(* IEC 61131-3 sources: Antarbhukti-LLM/DatasetCreation/SeedSTs/batch1_filtered_BASIC, 119 files *)

(* ---- A_TRIG.ST ---- *)
(*@PROPERTIES_EX@
TYPE: POU
LOCALE: 0
IEC_LANGUAGE: ST
PLC_TYPE: independent
PROC_TYPE: independent
GROUP: LOGIC.GENERATORS
*)
(*@KEY@:DESCRIPTION*)
version 1.1	23. oct. 2008
programmer 	hugo
tested by	oscat

this block is similar to the IEC Standard R_trig and F_trig but it monitors a REAL for change.
if the valiue on IN changes more then D from the last value it will generate trigger and display the difference in output D.
the trigger will only be active for one cycle.
(*@KEY@:END_DESCRIPTION*)
FUNCTION_BLOCK A_TRIG

(*Group:Default*)

VAR_INPUT
	IN :	REAL;
	RES :	REAL;
END_VAR

VAR_OUTPUT
	Q :	BOOL;
	D :	REAL;
END_VAR

VAR
	last_in :	REAL;
END_VAR

(*@KEY@: WORKSHEET
NAME: A_TRIG
IEC_LANGUAGE: ST
*)
D := IN - LAST_IN;
IF ABS(D) >= res THEN
	Q := TRUE;
	last_in := IN;
ELSE
	Q := FALSE;
END_IF;

(* revision history

hm 	16. jul. 2008	rev 1.0
	original version released

hm	23. oct. 2008	rev 1.1
	code optimization
*)
(*@KEY@: END_WORKSHEET *)
END_FUNCTION_BLOCK

(* ---- AIN1.ST ---- *)
(*@PROPERTIES_EX@
TYPE: POU
LOCALE: 0
IEC_LANGUAGE: ST
PLC_TYPE: independent
PROC_TYPE: independent
GROUP: ENGINEERING.SIGNAL_PROCESSING
*)
(*@KEY@:DESCRIPTION*)
version 1.3	10. mar. 2009
programmer 	oscat
tested by	tobias

Ain1 converts signals from A/D converters or other digital sources to an internal real value.

(*@KEY@:END_DESCRIPTION*)
FUNCTION_BLOCK AIN1

(*Group:Default*)

VAR_INPUT
	IN :	DWORD;
	SIGN_BIT :	INT := 255;
	ERROR_BIT :	INT := 255;
	ERROR_CODE_EN :	BOOL := FALSE;
	ERROR_CODE :	DWORD;
	OVERFLOW_BIT :	INT := 255;
	OVERFLOW_CODE_EN :	BOOL;
	OVERFLOW_CODE :	DWORD;
	BIT_0 :	INT;
	BIT_N :	INT := 31;
	OUT_MIN :	REAL;
	OUT_MAX :	REAL := 10.0;
	CODE_MIN :	DWORD;
	CODE_MAX :	DWORD := DWORD#16#FFFFFFFF;
	ERROR_OUTPUT :	REAL;
	OVERFLOW_OUTPUT :	REAL := 10.0;
END_VAR

VAR_OUTPUT
	OUT :	REAL;
	SIGN :	BOOL;
	ERROR :	BOOL;
	OVERFLOW :	BOOL;
END_VAR

VAR
	tB :	DWORD;
END_VAR

(*@KEY@: WORKSHEET
NAME: AIN1
IEC_LANGUAGE: ST
*)
(* extract error bit *)
error := ((SHR_DWORD(in,error_bit) AND DWORD#16#0000_0001) = DWORD#1) OR (error_code_en AND error_code = in);
IF error THEN
	out := error_output;
	RETURN;
END_IF;

(* strip off the data input *)
tb := SHR_DWORD(SHL_DWORD(in, 31 - bit_N), 31 - bit_N + Bit_0);

(* extract overflow bit *)
overflow := ((SHR_DWORD(in,overflow_bit) AND DWORD#16#0000_0001) = DWORD#1) OR (overflow_code_en AND overflow_code = in) OR (tb < code_min OR tb > code_max);
IF overflow THEN
	out := overflow_output;
	RETURN;
END_IF;

(* extract sign bit *)
sign := (SHR_DWORD(in,sign_bit) AND DWORD#16#0000_0001) = DWORD#1;

(* convert in to out *)
out := (UDINT_TO_REAL(DWORD_TO_UDINT(tb) - DWORD_TO_UDINT(code_min)) * (out_max - out_min) / UDINT_TO_REAL(DWORD_TO_UDINT(code_max) - DWORD_TO_UDINT(code_min)) + out_min);
IF sign THEN out := out * -1.0; END_IF;

(* revision history
hm	23. feb 2008	rev 1.0
	original version

hm	16. mar 2008	rev 1.1
	added type conversions to avoid warnngs under codesys 30

hm	22. apr. 2008	rev 1.2
	corrected error in formula when code_min was set
	corrected error when sign bit was used
	optimized code for better performance

hm	10. mar. 2009	rev 1.3
	real constants updated to new systax using dot

*)

(* extract error bit *)
error := ((SHR_DWORD(in,error_bit) AND DWORD#16#0000_0001) = DWORD#1) OR (error_code_en AND error_code = in);
IF error THEN
	out := error_output;
	RETURN;
END_IF;

(* strip off the data input *)
tb := SHR_DWORD(SHL_DWORD(in, 31 - bit_N), 31 - bit_N + Bit_0);

(* extract overflow bit *)
overflow := ((SHR_DWORD(in,overflow_bit) AND DWORD#16#0000_0001) = DWORD#1) OR (overflow_code_en AND overflow_code = in) OR (tb < code_min OR tb > code_max);
IF overflow THEN
	out := overflow_output;
	RETURN;
END_IF;

(* extract sign bit *)
sign := (SHR_DWORD(in,sign_bit) AND DWORD#16#0000_0001) = DWORD#1;

(* convert in to out *)
out := (UDINT_TO_REAL(DWORD_TO_UDINT(tb) - DWORD_TO_UDINT(code_min)) * (out_max - out_min) / UDINT_TO_REAL(DWORD_TO_UDINT(code_max) - DWORD_TO_UDINT(code_min)) + out_min);
IF sign THEN out := out * - 1.0; END_IF;

(* revision history
hm	23. feb 2008	rev 1.0
	original version

hm	16. mar 2008	rev 1.1
	added type conversions to avoid warnngs under codesys 30

hm	22. apr. 2008	rev 1.2
	corrected error in formula when code_min was set
	corrected error when sign bit was used
	optimized code for better performance

hm	10. mar. 2009	rev 1.3
	real constants updated to new systax using dot

*)

(*@KEY@: END_WORKSHEET *)
END_FUNCTION_BLOCK

(* ---- ALARM_2.ST ---- *)
(*@PROPERTIES_EX@
TYPE: POU
LOCALE: 0
IEC_LANGUAGE: ST
PLC_TYPE: independent
PROC_TYPE: independent
GROUP: ENGINEERING.MEASUREMENTS
*)
(*@KEY@:DESCRIPTION*)
version 1.1	11. mar. 2009
programmer 	hugo
tested BY	tobias

ALARM_2 will check two pairs of limits and signal when the input is above or below a set limit.
with the input HYS a hysteresis can be defined for all limits.
(*@KEY@:END_DESCRIPTION*)
FUNCTION_BLOCK ALARM_2

(*Group:Default*)

VAR_INPUT
	X :	REAL;
	LO_1 :	REAL;
	HI_1 :	REAL;
	LO_2 :	REAL;
	HI_2 :	REAL;
	HYS :	REAL;
END_VAR

VAR_OUTPUT
	Q1_LO :	BOOL;
	Q1_HI :	BOOL;
	Q2_LO :	BOOL;
	Q2_HI :	BOOL;
END_VAR

VAR
	tmp :	REAL;
END_VAR

(*@KEY@: WORKSHEET
NAME: ALARM_2
IEC_LANGUAGE: ST
*)
tmp := X - Hys * 0.5;
IF tmp > LO_1 THEN Q1_LO := FALSE; END_IF;
IF tmp > LO_2 THEN Q2_LO := FALSE; END_IF;
IF tmp > HI_1 THEN Q1_HI := TRUE; END_IF;
IF tmp > HI_2 THEN Q2_HI := TRUE; END_IF;
tmp := tmp + hys;
IF tmp < LO_1 THEN Q1_LO := TRUE; END_IF;
IF tmp < LO_2 THEN Q2_LO := TRUE; END_IF;
IF tmp < HI_1 THEN Q1_HI := FALSE; END_IF;
IF tmp < HI_2 THEN Q2_HI := FALSE; END_IF;

(* revision history
hm	19. may. 2008		rev 1.0
	original version

hm	11. mar. 2009	rev 1.1
	improved code
*)

(*@KEY@: END_WORKSHEET *)
END_FUNCTION_BLOCK

(* ---- B_TRIG.ST ---- *)
(*@PROPERTIES_EX@
TYPE: POU
LOCALE: 0
IEC_LANGUAGE: ST
PLC_TYPE: independent
PROC_TYPE: independent
GROUP: LOGIC.GENERATORS
*)
(*@KEY@:DESCRIPTION*)
version 1.0	4 aug 2006
programmer 	hugo
tested by	tobias

this block is similar to R_trig and F_trig but it generates a pulse on rising and falling edge.
(*@KEY@:END_DESCRIPTION*)
FUNCTION_BLOCK B_TRIG

(*Group:Default*)

VAR_INPUT
	CLK :	BOOL;
END_VAR

VAR_OUTPUT
	Q :	BOOL := FALSE;
END_VAR

VAR
	edge :	BOOL := FALSE;
END_VAR

(*@KEY@: WORKSHEET
NAME: B_TRIG
IEC_LANGUAGE: ST
*)
Q := clk XOR edge;
edge := CLK;
(*@KEY@: END_WORKSHEET *)
END_FUNCTION_BLOCK

(* ---- CALIBRATE.ST ---- *)
(*@PROPERTIES_EX@
TYPE: POU
LOCALE: 0
IEC_LANGUAGE: ST
PLC_TYPE: independent
PROC_TYPE: independent
GROUP: ENGINEERING.MEASUREMENTS
*)
(*@KEY@:DESCRIPTION*)
version 1.3	11. mar. 2009
programmer 	hugo
tested BY	hans

Calibrate allows for offset and scale calibration of an analog input.
offset is calibrated to a stored reference Y_offset while CO is true.
after the offset is calibrated, scale can be calibrated to a reference value Y_scale while CS is true.
*)
(*@KEY@:END_DESCRIPTION*)
FUNCTION_BLOCK CALIBRATE

(*Group:Default*)

VAR_INPUT
	X :	REAL;
	CO :	BOOL;
	CS :	BOOL;
	Y_OFFSET :	REAL;
	Y_SCALE :	REAL;
END_VAR

VAR_OUTPUT
	Y :	REAL;
END_VAR

VAR RETAIN
	offset :	REAL;
	Scale :	REAL := 1.0;
END_VAR

(*@KEY@: WORKSHEET
NAME: CALIBRATE
IEC_LANGUAGE: ST
*)
(* check for calibration *)
IF CO THEN
	OFFSET := Y_Offset - X;
ELSIF CS THEN
	SCALE := Y_scale / (X + OFFSET);
END_IF;
(* calculate output *)
Y := (X + OFFSET) * SCALE;

(* revision history
hm 22.2.2007		rev 1.2
	changed VAR RETAIN PERSISTENT to VAR RETAIN for better compatibility
	wago lon contollers do not support persisitent

hm	11. mar. 2009	rev 1.3
	changed real constants to use dot syntax

*)
(*@KEY@: END_WORKSHEET *)
END_FUNCTION_BLOCK

(* ---- CLICK_CNT.ST ---- *)
(*@PROPERTIES_EX@
TYPE: POU
LOCALE: 0
IEC_LANGUAGE: ST
PLC_TYPE: independent
PROC_TYPE: independent
GROUP: LOGIC.GENERATORS
*)
(*@KEY@:DESCRIPTION*)
version 1.0	16. jul. 2008
programmer 	hugo
tested by	oscat

this Module decodes a specified number of clicks.
the output trig is high for one cycle if N clicks are present within a specified time TC.
(*@KEY@:END_DESCRIPTION*)
FUNCTION_BLOCK CLICK_CNT

(*Group:Default*)

VAR_INPUT
	IN :	BOOL;
	N :	INT;
	TC :	TIME;
END_VAR

VAR_OUTPUT
	Q :	BOOL;
END_VAR

VAR
	tx :	TP;
	edge :	BOOL;
	cnt :	INT := INT#-1;
END_VAR

(*@KEY@: WORKSHEET
NAME: CLICK_CNT
IEC_LANGUAGE: ST
*)
(* Q shall only be active for one cycle only *)
Q := FALSE;

IF in AND NOT edge AND NOT tx.q THEN
	(* a rising edge on in sets the counter to 0 *)
	cnt := 0;
ELSIF tx.Q AND NOT IN AND edge THEN
	(* count falling edges when tp.q is true *)
	cnt := cnt + 1;
ELSIF NOT tx.Q THEN
	Q := cnt=N;
	cnt := -1;
END_IF;

(* remember the status of IN *)
edge := IN;
tx(in := IN, pt := TC);

(* revision history

hm 	16. jul. 2008	rev 1.0
	original version released

*)
(*@KEY@: END_WORKSHEET *)
END_FUNCTION_BLOCK

(* ---- CLICK_DEC.ST ---- *)
(*@PROPERTIES_EX@
TYPE: POU
LOCALE: 0
IEC_LANGUAGE: ST
PLC_TYPE: independent
PROC_TYPE: independent
GROUP: LOGIC.GENERATORS
*)
(*@KEY@:DESCRIPTION*)
version 1.1	14. mar. 2009
programmer 	hugo
tested by	oscat

this Module detects a rising edge on In and decodes the amount of falling edges (Pulses) within a specified time TC.
the outputs Q0..Q3 will go true for one cycle and the amount of clicks within a specified time TC.
if only a rising egde is detected within TC Q0 will respond, Q1 for 1 pulse and so on..

(*@KEY@:END_DESCRIPTION*)
FUNCTION_BLOCK CLICK_DEC

(*Group:Default*)

VAR_INPUT
	IN :	BOOL;
	TC :	TIME;
END_VAR

VAR_OUTPUT
	Q0 :	BOOL;
	Q1 :	BOOL;
	Q2 :	BOOL;
	Q3 :	BOOL;
END_VAR

VAR
	tx :	TP;
	edge :	BOOL;
	cnt :	INT := INT#-1;
END_VAR

(*@KEY@: WORKSHEET
NAME: CLICK_DEC
IEC_LANGUAGE: ST
*)
(* Q shall only be active for one cycle only *)
IF in = FALSE THEN
	Q0 := FALSE;
	Q1 := FALSE;
	Q2 := FALSE;
	Q3 := FALSE;
END_IF;

IF in AND NOT edge AND NOT tx.q THEN
	(* a rising edge on in sets the counter to 0 *)
	cnt := 0;
ELSIF tx.Q AND NOT IN AND edge THEN
	(* count falling edges when tp.q is true *)
	cnt := cnt + 1;
ELSIF NOT tx.Q THEN
	CASE cnt OF
		0 : Q0 := TRUE;
		1 : Q1 := TRUE;
		2 : Q2 := TRUE;
		3 : Q3 := TRUE;
	END_CASE;
	cnt := -1;
END_IF;

(* remember the status of IN *)
edge := IN;
tx(in := IN, pt := TC);

(* revision history

hm 17. jul. 2008	rev 1.0
	original version released

hm	14. mar. 2009	rev 1.1
	removed double assignments

*)
(*@KEY@: END_WORKSHEET *)
END_FUNCTION_BLOCK

(* ---- CLK_DIV.ST ---- *)
(*@PROPERTIES_EX@
TYPE: POU
LOCALE: 0
IEC_LANGUAGE: ST
PLC_TYPE: independent
PROC_TYPE: independent
GROUP: LOGIC.GENERATORS
*)
(*@KEY@:DESCRIPTION*)
version 1.1	2 jan 2008
programmer 	hugo
tested by	tobias

this is a clock divider
each output divides the signal by 2
Q0 = clk / 2 , Q1 = Q0 / 2 and so on.
the outputs have a 50% duty cycle each.
(*@KEY@:END_DESCRIPTION*)
FUNCTION_BLOCK CLK_DIV

(*Group:Default*)

VAR_INPUT
	CLK :	BOOL;
	RST :	BOOL;
END_VAR

VAR_OUTPUT
	Q0 :	BOOL := FALSE;
	Q1 :	BOOL := FALSE;
	Q2 :	BOOL := FALSE;
	Q3 :	BOOL := FALSE;
	Q4 :	BOOL := FALSE;
	Q5 :	BOOL := FALSE;
	Q6 :	BOOL := FALSE;
	Q7 :	BOOL := FALSE;
END_VAR

VAR
	cnt :	BYTE := 0;
END_VAR

(*@KEY@: WORKSHEET
NAME: CLK_DIV
IEC_LANGUAGE: ST
*)
IF rst THEN
	cnt:= BYTE#0;
	Q0 := FALSE;
	Q1 := FALSE;
	Q2 := FALSE;
	Q3 := FALSE;
	Q4 := FALSE;
	Q5 := FALSE;
	Q6 := FALSE;
	Q7 := FALSE;
ELSIF clk THEN
	cnt:= USINT_TO_BYTE(BYTE_TO_USINT(cnt) + USINT#1);

    Q0 := BIT_OF_DWORD(BYTE_TO_DWORD(cnt),0); (* Q0 := cnt.X0; *)
    Q1 := BIT_OF_DWORD(BYTE_TO_DWORD(cnt),1); (* Q1 := cnt.X1; *)
    Q2 := BIT_OF_DWORD(BYTE_TO_DWORD(cnt),2); (* Q2 := cnt.X2; *)
    Q3 := BIT_OF_DWORD(BYTE_TO_DWORD(cnt),3); (* Q3 := cnt.X3; *)
    Q4 := BIT_OF_DWORD(BYTE_TO_DWORD(cnt),4); (* Q4 := cnt.X4; *)
    Q5 := BIT_OF_DWORD(BYTE_TO_DWORD(cnt),5); (* Q5 := cnt.X5; *)
    Q6 := BIT_OF_DWORD(BYTE_TO_DWORD(cnt),6); (* Q6 := cnt.X6; *)
    Q7 := BIT_OF_DWORD(BYTE_TO_DWORD(cnt),7); (* Q7 := cnt.X7; *)

END_IF;

(* revision history
hm	4. aug. 2006	rev 1.0
	original version

hm	2. jan 2008		rev 1.1
	improved performance

*)
(*@KEY@: END_WORKSHEET *)
END_FUNCTION_BLOCK

(* ---- CLK_N.ST ---- *)
(*@PROPERTIES_EX@
TYPE: POU
LOCALE: 0
IEC_LANGUAGE: ST
PLC_TYPE: independent
PROC_TYPE: independent
GROUP: LOGIC.GENERATORS
*)
(*@KEY@:DESCRIPTION*)
version 1.0	17 sep 2007
programmer 	hugo
tested by	tobias

clk_N uses the internal sps time to generate one pulse every N ms
every pulse is only valid for one cycle so that a edge trigger is not necessary
clk_gen generates pulses depending on the accuracy of the system clock.
The input N controlls the period time of the clock.
N=0 equals 2ms, N=1 equals 4ms, N=2 equals 8ms, N=3 equals 16ms ....

be careful, 1ms clocks will only work on very powerful sps cpu's
(*@KEY@:END_DESCRIPTION*)
FUNCTION_BLOCK CLK_N

(*Group:Default*)

VAR_INPUT
	N :	INT;
END_VAR

VAR_OUTPUT
	Q :	BOOL;
END_VAR

VAR
	T_PLC_MS :	T_PLC_MS;
	edge :	BOOL;
	clk :	BOOL;
END_VAR

(*@KEY@: WORKSHEET
NAME: CLK_N
IEC_LANGUAGE: ST
*)
T_PLC_MS();
clk := BIT_OF_DWORD(SHR(UDINT_TO_DWORD(T_PLC_MS.T_PLC_MS),N),0);
Q := clk XOR edge;
edge := clk;

(* revision history
hm	16. dec 2007		rev 1.0
	original version

*)
(*@KEY@: END_WORKSHEET *)
END_FUNCTION_BLOCK

(* ---- CLK_PRG.ST ---- *)
(*@PROPERTIES_EX@
TYPE: POU
LOCALE: 0
IEC_LANGUAGE: ST
PLC_TYPE: independent
PROC_TYPE: independent
GROUP: LOGIC.GENERATORS
*)
(*@KEY@:DESCRIPTION*)
version 1.3	25. oct. 2008
programmer 	hugo
tested by	tobias

clk_prg uses the internal sps time to generate a clock with programmable period time.
the period time is defined for 10ms .. 65s
the first cycle after start is a clk pulse and then depending on the programmed period time a delay.
every pulse is only valid for one cycle.
the accuracy of clk_prg is depending on the accuracy of the system clock.
(*@KEY@:END_DESCRIPTION*)
FUNCTION_BLOCK CLK_PRG

(*Group:Default*)

VAR_INPUT
	PT :	TIME := T#10ms;
END_VAR

VAR_OUTPUT
	Q :	BOOL;
END_VAR

VAR
	init :	BOOL := FALSE;
	last :	TIME;
	tx :	TIME;
	T_PLC_MS :	T_PLC_MS;
END_VAR

(*@KEY@: WORKSHEET
NAME: CLK_PRG
IEC_LANGUAGE: ST
*)
(* read system time *)
T_PLC_MS();
tx:= UDINT_TO_TIME(T_PLC_MS.T_PLC_MS);

(* initialize on startup *)
IF NOT init THEN
	init := TRUE;
	last := tx - pt;
END_IF;

(* generate output pulse when next_pulse is reached *)
Q := tx - last >= pt;
IF Q THEN last := tx; END_IF;

(* revision hiostory

hm 25 feb 2007	rev 1.1
	rewritten code for higher performance
	pt can now be changed during runtime

hm	17. sep 2007	rev 1.2
	replaced time() with t_plc_ms() for compatibility reasons

hm	25. oct. 2008	rev 1.3
	optimized code

*)
(*@KEY@: END_WORKSHEET *)
END_FUNCTION_BLOCK

(* ---- CLK_PULSE.ST ---- *)
(*@PROPERTIES_EX@
TYPE: POU
LOCALE: 0
IEC_LANGUAGE: ST
PLC_TYPE: independent
PROC_TYPE: independent
GROUP: LOGIC.GENERATORS
*)
(*@KEY@:DESCRIPTION*)
version 1.2		16 feb 2011
programmer 	    hugo
tested by		oscat

clk_pulse uses the internal sps time to generate a clock with programmable period time.
the period time is defined for 10ms .. 65s.
pulse generation is continuous if N = 0 and for n pulses otherwise.
the first cycle after start is a clk pulse and then depending on the programmed period time a delay.
every pulse is only valid for one cycle so that a edge trigger is not necessary
clk_prg depending on the accuracy of the system clock.

(*@KEY@:END_DESCRIPTION*)
FUNCTION_BLOCK CLK_PULSE

(*Group:Default*)

VAR_INPUT
	PT :	TIME;
	N :	INT;
	RST :	BOOL;
END_VAR

VAR_OUTPUT
	Q :	BOOL;
	CNT :	INT;
	RUN :	BOOL;
END_VAR

VAR
	tx :	UDINT;
	tn :	UDINT;
	init :	BOOL;
	T_PLC_MS :	T_PLC_MS;
END_VAR

(*@KEY@: WORKSHEET
NAME: CLK_PULSE
IEC_LANGUAGE: ST
*)
(* read system *)
T_PLC_MS();
tx:= T_PLC_MS.T_PLC_MS;
Q := FALSE;				(* reset Q we generate pulses only for one cycle *)
RUN := CNT < N;

IF NOT init OR RST THEN
	init := TRUE;
	CNT := 0;
	tn := tx - TIME_TO_UDINT(PT);
	RUN := FALSE;
ELSIF (cnt < N OR N = 0) AND tx - tn >= TIME_TO_UDINT(PT) THEN		(* generate a pulse *)
	CNT := CNT + 1;
	Q := TRUE;
	tn := tn + TIME_TO_UDINT(PT);
END_IF;

(* revision history
hm		4. aug 2006		rev 1.0
	original version

hm		17. sep 2007	rev 1.1
	replaced time() with T_PLC_S() for compatblity reasons

hm		16. feb. 2011	rev 1.2
	fixed an error when timer overflows
*)
(*@KEY@: END_WORKSHEET *)
END_FUNCTION_BLOCK

(* ---- CONTROL_SET1.ST ---- *)
(*@PROPERTIES_EX@
TYPE: POU
LOCALE: 0
IEC_LANGUAGE: ST
PLC_TYPE: independent
PROC_TYPE: independent
GROUP: ENGINEERING.CONTROL
*)
(*@KEY@:DESCRIPTION*)
version 1.1	11. mar. 2009
programmer 	hugo
tested by	tobias

takahashi calculates controller parameters for P, PI and PID controllers based on the ziegler nichols method.

(*@KEY@:END_DESCRIPTION*)
FUNCTION_BLOCK CONTROL_SET1

(*Group:Default*)

VAR_INPUT
	KT :	REAL;
	TT :	REAL;
	PI :	BOOL;
	PID :	BOOL;
	P_K :	REAL := 0.5;
	PI_K :	REAL := 0.45;
	PI_TN :	REAL := 0.83;
	PID_K :	REAL := 0.6;
	PID_TN :	REAL := 0.5;
	PID_TV :	REAL := 0.125;
END_VAR

VAR_OUTPUT
	KP :	REAL;
	TN :	REAL;
	TV :	REAL;
	KI :	REAL;
	KD :	REAL;
END_VAR

(*@KEY@: WORKSHEET
NAME: CONTROL_SET1
IEC_LANGUAGE: ST
*)
IF pi AND PID THEN
	KP := 0.0;
	TN := 0.0;
	TV := 0.0;
ELSIF PID THEN
	KP := PID_K * Kt;
	TN := PID_TN * Tt;
	TV := PID_TV * Tt;
ELSIF PI THEN
	KP := PI_K * Kt;
	TN := PI_TN * Tt;
ELSE
	KP := P_K * Kt;
END_IF;

(* KI and KD are calculated *)
IF tn > 0.0 THEN KI := KP / TN; ELSE KI := 0.0; END_IF;
KD := KP * TV;

(* revision history
hm	4. nov 2007	rev 1.0
	original version

hm	11. mar. 2009	rev 1.1
	real constants updated to new systax using dot

*)
(*@KEY@: END_WORKSHEET *)
END_FUNCTION_BLOCK

(* ---- CONTROL_SET2.ST ---- *)
(*@PROPERTIES_EX@
TYPE: POU
LOCALE: 0
IEC_LANGUAGE: ST
PLC_TYPE: independent
PROC_TYPE: independent
GROUP: ENGINEERING.CONTROL
*)
(*@KEY@:DESCRIPTION*)
version 1.1	11. mar. 2009
programmer 	hugo
tested by	tobias

takahashi calculates controller parameters for P, PI and PID controllers based on the ziegler nichols method.

(*@KEY@:END_DESCRIPTION*)
FUNCTION_BLOCK CONTROL_SET2

(*Group:Default*)

VAR_INPUT
	KS :	REAL;
	TU :	REAL;
	TG :	REAL;
	PI :	BOOL;
	PID :	BOOL;
	P_K :	REAL := 1.0;
	PI_K :	REAL := 0.9;
	PI_TN :	REAL := 3.33;
	PID_K :	REAL := 1.2;
	PID_TN :	REAL := 2.0;
	PID_TV :	REAL := 0.5;
END_VAR

VAR_OUTPUT
	KP :	REAL;
	TN :	REAL;
	TV :	REAL;
	KI :	REAL;
	KD :	REAL;
END_VAR

VAR
	TX :	REAL;
END_VAR

(*@KEY@: WORKSHEET
NAME: CONTROL_SET2
IEC_LANGUAGE: ST
*)
IF TU > 0.0 AND KS > 0.0 THEN TX := TG / TU / KS; END_IF;
IF pi AND PID THEN
	KP := 0.0;
	TN := 0.0;
	TV := 0.0;
ELSIF PID THEN
	KP := PID_K * TX;
	TN := PID_TN * TU;
	TV := PID_TV * TU;
ELSIF PI THEN
	KP := PI_K * TX;
	TN := PI_TN * TU;
ELSE
	KP := P_K * TX;
END_IF;

(* KI and KD are calculated *)
IF TN > 0.0 THEN KI := KP / TN; ELSE KI := 0.0; END_IF;
KD := KP * TV;

(* revision history
hm	4. nov 2007	rev 1.0
	original version

hm	11. mar. 2009	rev 1.1
	real constants updated to new systax using dot

*)
(*@KEY@: END_WORKSHEET *)
END_FUNCTION_BLOCK

(* ---- COUNT_BR.ST ---- *)
(*@PROPERTIES_EX@
TYPE: POU
LOCALE: 0
IEC_LANGUAGE: ST
PLC_TYPE: independent
PROC_TYPE: independent
GROUP: LOGIC.FF_EDGE_TRIGGERED
*)
(*@KEY@:DESCRIPTION*)
version 1.0	16 jan 2008
programmer 	hugo
tested BY	tobias

Count_R is a byte counter with independen up and dn inputs. the counter counts from 0 to mx and continues at 0 after is has reached mx
a step input sets the counters stepping width.
(*@KEY@:END_DESCRIPTION*)
FUNCTION_BLOCK COUNT_BR

(*Group:Default*)

VAR_INPUT
	SET :	BOOL;
	IN :	BYTE;
	UP :	BOOL;
	DN :	BOOL;
	STEP :	BYTE := BYTE#1;
	MX :	BYTE := BYTE#255;
	RST :	BOOL;
END_VAR

VAR_OUTPUT
	CNT :	BYTE;
END_VAR

VAR
	last_up :	BOOL;
	last_dn :	BOOL;
END_VAR

(*@KEY@: WORKSHEET
NAME: COUNT_BR
IEC_LANGUAGE: ST
*)
IF rst THEN
	cnt := BYTE#0;
ELSIF set THEN
	cnt := INT_TO_BYTE(LIMIT(0,_BYTE_TO_INT(in),_BYTE_TO_INT(mx)));
ELSIF up AND NOT last_up THEN
	cnt := INT_TO_BYTE(inc(_BYTE_TO_INT(cnt),_BYTE_TO_INT(step),_BYTE_TO_INT(mx)));
ELSIF dn AND NOT last_dn THEN
	cnt := INT_TO_BYTE(inc(_BYTE_TO_INT(cnt),_BYTE_TO_INT(step) * -1,_BYTE_TO_INT(mx)));
END_IF;
last_up := up;
last_dn := dn;

(* revision history
hm	16. jan 2008	rev 1.0
	original version

*)
(*@KEY@: END_WORKSHEET *)
END_FUNCTION_BLOCK

(* ---- COUNT_DR.ST ---- *)
(*@PROPERTIES_EX@
TYPE: POU
LOCALE: 0
IEC_LANGUAGE: ST
PLC_TYPE: independent
PROC_TYPE: independent
GROUP: LOGIC.FF_EDGE_TRIGGERED
*)
(*@KEY@:DESCRIPTION*)
version 1.1	20. jan. 2011
programmer 	hugo
tested BY	tobias

Count_DR is a DWORD counter with independen up and dn inputs. the counter counts from 0 to mx and continues at 0 after is has reached mx
a step input sets the counters stepping width.
(*@KEY@:END_DESCRIPTION*)
FUNCTION_BLOCK COUNT_DR

(*Group:Default*)

VAR_INPUT
	SET :	BOOL;
	IN :	DWORD;
	UP :	BOOL;
	DN :	BOOL;
	STEP :	DWORD := DWORD#1;
	MX :	DWORD := DWORD#16#FFFF_FFFF;
	RST :	BOOL;
END_VAR

VAR_OUTPUT
	CNT :	DWORD;
END_VAR

VAR
	CNT2 :	UDINT;
	STEP2 :	UDINT;
	MX2 :	UDINT;
	last_up :	BOOL;
	last_dn :	BOOL;
END_VAR

(*@KEY@: WORKSHEET
NAME: COUNT_DR
IEC_LANGUAGE: ST
*)
STEP2 := DWORD_TO_UDINT(STEP);
MX2   := DWORD_TO_UDINT(MX);
CNT2  := DWORD_TO_UDINT(CNT);

IF rst THEN
	CNT2 := UDINT#0;
ELSIF set THEN
	CNT2 := LIMIT(UDINT#0,DWORD_TO_UDINT(in),mx2);
ELSIF up AND NOT last_up THEN
	IF STEP2 > MX2 - CNT2 THEN
		CNT2 := CNT2 - MX2 + STEP2 - UDINT#1;
	ELSE
		CNT2 := CNT2 + STEP2;
	END_IF;
ELSIF dn AND NOT last_dn THEN
	IF STEP2 > CNT2 THEN
		CNT2 := CNT2 - STEP2 + MX2 + UDINT#1;
	ELSE
		CNT2 := CNT2 - STEP2;
	END_IF;
END_IF;
last_up := up;
last_dn := dn;

CNT := UDINT_TO_DWORD(CNT2);

(* revision history
hm	12. jun 2008	rev 1.0
	original version

hm	20. jan. 2011	rev 1.1
	corrected init value of MX to 16#FFFFFFFF

*)
(*@KEY@: END_WORKSHEET *)
END_FUNCTION_BLOCK

(* ---- CTRL_OUT.ST ---- *)
(*@PROPERTIES_EX@
TYPE: POU
LOCALE: 0
IEC_LANGUAGE: ST
PLC_TYPE: independent
PROC_TYPE: independent
GROUP: ENGINEERING.CONTROL
*)
(*@KEY@:DESCRIPTION*)
version 1.1	3. nov 2008
programmer 	hugo
tested by	oscat
(*@KEY@:END_DESCRIPTION*)
FUNCTION_BLOCK CTRL_OUT

(*Group:Default*)

VAR_INPUT
	CI :	REAL;
	OFFSET :	REAL;
	MAN_IN :	REAL;
	LIM_L :	REAL;
	LIM_H :	REAL;
	MANUAL :	BOOL;
END_VAR

VAR_OUTPUT
	Y :	REAL;
	LIM :	BOOL;
END_VAR

(*@KEY@: WORKSHEET
NAME: CTRL_OUT
IEC_LANGUAGE: ST
*)
Y := SEL(manual, CI, MAN_IN) + OFFSET;

(* Limit the output *)
IF Y >= LIM_H THEN
	Y := LIM_H;
	LIM := TRUE;
ELSIF Y <= lim_L THEN
	Y := LIM_L;
	LIM := TRUE;
ELSE
	LIM := FALSE;
END_IF;

(* revision history
hm 	2. jun. 2008 	rev 1.0
	original version

hm	3. nov. 2008	rev 1.1
	optimized code
*)
(*@KEY@: END_WORKSHEET *)
END_FUNCTION_BLOCK

(* ---- CTRL_PI.ST ---- *)
(*@PROPERTIES_EX@
TYPE: POU
LOCALE: 0
IEC_LANGUAGE: ST
PLC_TYPE: independent
PROC_TYPE: independent
GROUP: ENGINEERING.CONTROL
*)
(*@KEY@:DESCRIPTION*)
version 2.0	30. jun. 2008
programmer 	hugo
tested by	oscat

FT_PI is a PI controller with manual functionality.
The PID controller works according to the fomula Y = e *(KP+ KI * INTEG(e) ) + offset, while e = set_point - actual.
a rst will reset all internal data, while a switch to manual will cause the controller to follow the function Y = manual_in + offset.
limit_h and Limit_l set the possible output range of Y.
the output flags lim will signal that the output limits are active and overflow will signal that the integrator has reached its limits.

since rev 1.1 the "trapezregel is used for more accuracy.
rev 1.2 added selective integratin which means the integrative component is only active within a small range of the target value
this avoids the integrator to go to limits while an input setpoint change happened and is only causing overshoots.
the int_band is by default 100 which means the int is active all the time and if set to for example to 0.1 the integrator is only active
while the input is between 0.9 and 1.1 of the set_point value.

default values for KP = 1, TN = 1, TV = 1, LIMIT_L = -1000, LIMIT_H = +1000.
(*@KEY@:END_DESCRIPTION*)
FUNCTION_BLOCK CTRL_PI

(*Group:Default*)

VAR_INPUT
	ACT :	REAL;
	SET :	REAL;
	SUP :	REAL;
	OFS :	REAL;
	M_I :	REAL;
	MAN :	BOOL;
	RST :	BOOL := FALSE;
	KP :	REAL := 1.0;
	KI :	REAL := 1.0;
	LL :	REAL := -1000.0;
	LH :	REAL := 1000.0;
END_VAR

VAR_OUTPUT
	Y :	REAL;
	DIFF :	REAL;
	LIM :	BOOL;
END_VAR

VAR
	pi :	FT_PIWL;
	co :	CTRL_OUT;
END_VAR

(*@KEY@: WORKSHEET
NAME: CTRL_PI
IEC_LANGUAGE: ST
*)
DIFF := CTRL_IN(SET, ACT, SUP);
pi(in := DIFF, kp := KP, ki := KI, lim_l := LL, lim_h := LH, rst := RST);
co(ci := pi.Y, OFFSET := OFS, man_in := M_I, lim_l := LL, lim_h := LH, manual := MAN);
Y := co.Y;
LIM := co.LIM;

(* revision history
hm 	31.10.2007 	rev 1.0
	original version

hm	3.11.2007	rev 1.1
	added noise input to filter noise
	added output diff
	set limit output false when output is within limits
	overfolw was not set correctly

hm	5. jan 2008	rev 1.2
	improved performance

hm	30. jun. 2008	rev 2.0
	rewritten using new modular approach*)
(*@KEY@: END_WORKSHEET *)
END_FUNCTION_BLOCK

(* ---- CTRL_PID.ST ---- *)
(*@PROPERTIES_EX@
TYPE: POU
LOCALE: 0
IEC_LANGUAGE: ST
PLC_TYPE: independent
PROC_TYPE: independent
GROUP: ENGINEERING.CONTROL
*)
(*@KEY@:DESCRIPTION*)
version 2.0	30. jun. 2008
programmer 	hugo
tested by	oscat

FT_PI is a PI controller with manual functionality.
The PID controller works according to the fomula Y = e *(KP+ KI * INTEG(e) ) + offset, while e = set_point - actual.
a rst will reset all internal data, while a switch to manual will cause the controller to follow the function Y = manual_in + offset.
limit_h and Limit_l set the possible output range of Y.
the output flags lim will signal that the output limits are active.
(*@KEY@:END_DESCRIPTION*)
FUNCTION_BLOCK CTRL_PID

(*Group:Default*)

VAR_INPUT
	ACT :	REAL;
	SET :	REAL;
	SUP :	REAL;
	OFS :	REAL;
	M_I :	REAL;
	MAN :	BOOL;
	RST :	BOOL := FALSE;
	KP :	REAL := 1.0;
	TN :	REAL := 1.0;
	TV :	REAL := 1.0;
	LL :	REAL := -1000.0;
	LH :	REAL := 1000.0;
END_VAR

VAR_OUTPUT
	Y :	REAL;
	DIFF :	REAL;
	LIM :	BOOL;
END_VAR

VAR
	pid :	FT_PIDWL;
	co :	CTRL_OUT;
END_VAR

(*@KEY@: WORKSHEET
NAME: CTRL_PID
IEC_LANGUAGE: ST
*)
DIFF := CTRL_IN(SET, ACT, SUP);
pid(in := DIFF, kp := KP, tn := TN, tv := TV, lim_l := LL, lim_h := LH, rst := RST);
co(ci := pid.Y, OFFSET := OFS, man_in := M_I, lim_l := LL, lim_h := LH, manual := MAN);
Y := co.Y;
LIM := co.LIM;

(* revision history
hm 	31.10.2007 		rev 1.0
	original version

hm	3.11.2007		rev 1.1
	added noise input to filter noise
	added output diff
	set limit output false when output is within limits
	overfolw was not set correctly

hm	5. jan 2008		rev 1.2
	improved performance

hm	30. jun. 2008	rev 2.0
	rewritten using new modular approach

*)
(*@KEY@: END_WORKSHEET *)
END_FUNCTION_BLOCK

(* ---- CTRL_PWM.ST ---- *)
(*@PROPERTIES_EX@
TYPE: POU
LOCALE: 0
IEC_LANGUAGE: ST
PLC_TYPE: independent
PROC_TYPE: independent
GROUP: ENGINEERING.CONTROL
*)
(*@KEY@:DESCRIPTION*)
version 1.1	21. oct. 2008
programmer 	hugo
tested by	oscat
(*@KEY@:END_DESCRIPTION*)
FUNCTION_BLOCK CTRL_PWM

(*Group:Default*)

VAR_INPUT
	CI :	REAL;
	MAN_IN :	REAL;
	MANUAL :	BOOL;
	F :	REAL;
END_VAR

VAR_OUTPUT
	Q :	BOOL;
END_VAR

VAR
	PW :	PWM_DC;
END_VAR

(*@KEY@: WORKSHEET
NAME: CTRL_PWM
IEC_LANGUAGE: ST
*)
PW(F := F, DC := SEL(MANUAL,CI,MAN_IN));
Q := PW.Q;

(* revision history
hm 	3. jun. 2008 	rev 1.0
	original version

hm	21. oct. 2008	rev 1.1
	optimized code
*)
(*@KEY@: END_WORKSHEET *)
END_FUNCTION_BLOCK

(* ---- CYCLE_4.ST ---- *)
(*@PROPERTIES_EX@
TYPE: POU
LOCALE: 0
IEC_LANGUAGE: ST
PLC_TYPE: independent
PROC_TYPE: independent
GROUP: LOGIC.GENERATORS
*)
(*@KEY@:DESCRIPTION*)
version 1.0
programmer 	hugo
tested by	oscat
(*@KEY@:END_DESCRIPTION*)
FUNCTION_BLOCK CYCLE_4

(*Group:Default*)

VAR_INPUT
	E :	BOOL := TRUE;
	T0 :	TIME;
	T1 :	TIME;
	T2 :	TIME;
	T3 :	TIME;
	S0 :	BOOL;
	SX :	INT;
	SL :	BOOL;
END_VAR

VAR_OUTPUT
	STATE :	INT;
END_VAR

VAR
	tx :	TIME;
	last :	TIME;
	init :	BOOL;
	T_PLC_MS :	T_PLC_MS;
END_VAR

(*@KEY@: WORKSHEET
NAME: CYCLE_4
IEC_LANGUAGE: ST
*)
(* read system *)
T_PLC_MS();
tx:= UDINT_TO_TIME(T_PLC_MS.T_PLC_MS);

(* init on first cycle *)
IF NOT init THEN
	init := TRUE;
	last := tx;
END_IF;

IF E THEN
	IF SL THEN
		(* when sx > 0 then the state sx is forced to start *)
		state:= LIMIT(0,SX,3);
		last := tx;
		(* this is to avoid to reset sx from the calling programm it does work fine on codesys but i am not sure about other systems, because we are writing to an input *)
		SL := FALSE;
	ELSE
		CASE state OF
			0 :	(* wait for T0 and switch to next cycle *)
				IF tx - last >= T0 THEN
					state := 1;
					last := tx;
				END_IF;
			1 : (* wait for T1 over 1st cycle *)
				IF tx - last >= T1 THEN
					state := 2;
					last := tx;
				END_IF;
			2 : (* wait for T1 over 1st cycle *)
				IF tx - last >= T2 THEN
					state := 3;
					last := tx;
				END_IF;
			3 : (* wait for T2 over 2nd cycle *)
				IF tx - last >= T3 THEN
					IF S0 THEN State := 0; END_IF; (* if S0 is false, the sequence stops at state 3 *)
					last := tx;
				END_IF;
		END_CASE;
	END_IF;
ELSE
	state := 0;
	last := tx;
END_IF;

(*
hm	3. nov. 2008	rev 1.0
	original version

*)
(*@KEY@: END_WORKSHEET *)
END_FUNCTION_BLOCK

(* ---- D_TRIG.ST ---- *)
(*@PROPERTIES_EX@
TYPE: POU
LOCALE: 0
IEC_LANGUAGE: ST
PLC_TYPE: independent
PROC_TYPE: independent
GROUP: LOGIC.GENERATORS
*)
(*@KEY@:DESCRIPTION*)
version 1.1	19. feb 2008
programmer 	hugo
tested by	tobias

this block is similar to the IEC Standard R_trig and F_trig but it monitors a DWORD, WORD or Byte Variable instead and generated an Output Pulse for one cycle only when the input has changed.
an additional output x (Dword) will state the chage of the input.
Example: the input has chaged from 0001 to 0010 then the output x will be 2.
(*@KEY@:END_DESCRIPTION*)
FUNCTION_BLOCK D_TRIG

(*Group:Default*)

VAR_INPUT
	IN :	DWORD;
END_VAR

VAR_OUTPUT
	Q :	BOOL;
	X :	DWORD;
END_VAR

VAR
	last_in :	DWORD;
END_VAR

(*@KEY@: WORKSHEET
NAME: D_TRIG
IEC_LANGUAGE: ST
*)
Q := in <> last_in;
X := UDINT_TO_DWORD(DWORD_TO_UDINT(in) - DWORD_TO_UDINT(last_in));
last_in := in;

(* revision history

hm 	4.09.2007		rev 1.0
	original version released

hm	19. feb. 2008	rev 1.1
	performance improvement
*)
(*@KEY@: END_WORKSHEET *)
END_FUNCTION_BLOCK

(* ---- DEC_2.ST ---- *)
(*@PROPERTIES_EX@
TYPE: POU
LOCALE: 0
IEC_LANGUAGE: ST
PLC_TYPE: independent
PROC_TYPE: independent
GROUP: LOGIC.GATE_LOGIC
*)
(*@KEY@:DESCRIPTION*)
version 1.1	3 Mar 2007
programmer 	hugo
tested by	tobias

a bit input will be decoded to the two outputs Q0 or Q1
dependent on the value of A
A=0 decodes to Q0 and A=1 decodes to Q1
(*@KEY@:END_DESCRIPTION*)
FUNCTION_BLOCK DEC_2

(*Group:Default*)

VAR_INPUT
	D :	BOOL;
	A :	BOOL;
END_VAR

VAR_OUTPUT
	Q0 :	BOOL;
	Q1 :	BOOL;
END_VAR

(*@KEY@: WORKSHEET
NAME: DEC_2
IEC_LANGUAGE: ST
*)
Q0 := D AND NOT A;
Q1 := D AND A;

(* revision history
hm 3.3.2007	rev 1.1
	rewritten in ST for better compatibility
*)
(*@KEY@: END_WORKSHEET *)
END_FUNCTION_BLOCK

(* ---- DEC_4.ST ---- *)
(*@PROPERTIES_EX@
TYPE: POU
LOCALE: 0
IEC_LANGUAGE: ST
PLC_TYPE: independent
PROC_TYPE: independent
GROUP: LOGIC.GATE_LOGIC
*)
(*@KEY@:DESCRIPTION*)
version 1.1	3 Mar 2007
programmer 	hugo
tested by	tobias

a bit input will be decoded to one of the 4 outputs
dependent on the Adress on A0 and A1
(*@KEY@:END_DESCRIPTION*)
FUNCTION_BLOCK DEC_4

(*Group:Default*)

VAR_INPUT
	D :	BOOL;
	A0 :	BOOL;
	A1 :	BOOL;
END_VAR

VAR_OUTPUT
	Q0 :	BOOL;
	Q1 :	BOOL;
	Q2 :	BOOL;
	Q3 :	BOOL;
END_VAR

(*@KEY@: WORKSHEET
NAME: DEC_4
IEC_LANGUAGE: ST
*)
Q0 := D AND NOT A0 AND NOT A1;
Q1 := D AND A0 AND NOT A1;
Q2 := D AND NOT A0 AND A1;
Q3 := D AND A0 AND A1;

(* revision history
hm 3.3.2007	rev 1.1
	rewritten in ST for better compatibility

*)
(*@KEY@: END_WORKSHEET *)
END_FUNCTION_BLOCK

(* ---- DEC_8.ST ---- *)
(*@PROPERTIES_EX@
TYPE: POU
LOCALE: 0
IEC_LANGUAGE: ST
PLC_TYPE: independent
PROC_TYPE: independent
GROUP: LOGIC.GATE_LOGIC
*)
(*@KEY@:DESCRIPTION*)
version 1.3	28. mar. 2009
programmer 	hugo
tested by	oscat

a bit input will be decoded to one of the 8 outputs
dependent on the Adress on A0, A1 and A2

(*@KEY@:END_DESCRIPTION*)
FUNCTION_BLOCK DEC_8

(*Group:Default*)

VAR_INPUT
	D :	BOOL;
	A0 :	BOOL;
	A1 :	BOOL;
	A2 :	BOOL;
END_VAR

VAR_OUTPUT
	Q0 :	BOOL;
	Q1 :	BOOL;
	Q2 :	BOOL;
	Q3 :	BOOL;
	Q4 :	BOOL;
	Q5 :	BOOL;
	Q6 :	BOOL;
	Q7 :	BOOL;
END_VAR

VAR
	X :	BYTE;
END_VAR

(*@KEY@: WORKSHEET
NAME: DEC_8
IEC_LANGUAGE: ST
*)
X:=BIT_LOAD_B(X,A0,0); (* X.0 := A0; *)
X:=BIT_LOAD_B(X,A1,1); (* X.1 := A1; *)
X:=BIT_LOAD_B(X,A2,2); (* X.2 := A2; *)

Q0 := FALSE;
Q1 := FALSE;
Q2 := FALSE;
Q3 := FALSE;
Q4 := FALSE;
Q5 := FALSE;
Q6 := FALSE;
Q7 := FALSE;

CASE _BYTE_TO_INT(X) OF
	0 : Q0 := D;
	1 : Q1 := D;
	2 : Q2 := D;
	3 : Q3 := D;
	4 : Q4 := D;
	5 : Q5 := D;
	6 : Q6 := D;
	7 : Q7 := D;
END_CASE;

(* revision history
hm 3. mar. 2007	rev 1.1
	rewritten in ST for better compatibility

hm	26. oct. 2008	rev 1.2
	code optimized

hm	28. mar. 2009	rev 1.3
	replaced multiple assignments
*)
(*@KEY@: END_WORKSHEET *)
END_FUNCTION_BLOCK

(* ---- DELAY.ST ---- *)
(*@PROPERTIES_EX@
TYPE: POU
LOCALE: 0
IEC_LANGUAGE: ST
PLC_TYPE: independent
PROC_TYPE: independent
GROUP: ENGINEERING.SIGNAL_PROCESSING
*)
(*@KEY@:DESCRIPTION*)
version 1.5	23. mar. 2009
programmer 	hugo
tested by	oscat

this function block delays input values by each programm cycle
after N+1 cycles the in value has shifted to the out.
N can be any alue from 0 .. 32
if n = 0 the input will be present on the output without a delay.
f N > 32 then the output will be delayed by 32 cycles.
any high on rst will load the buffer with in.

(*@KEY@:END_DESCRIPTION*)
FUNCTION_BLOCK DELAY

(*Group:Default*)

VAR_INPUT
	IN :	REAL;
	N :	INT;
	RST :	BOOL;
END_VAR

VAR_OUTPUT
	OUT :	REAL;
END_VAR

VAR
	buf :	oscat_delay_buf;
	i :	INT;
	init :	BOOL;
	stop :	INT;
END_VAR

(*@KEY@: WORKSHEET
NAME: DELAY
IEC_LANGUAGE: ST
*)
stop := LIMIT(0,N,32) - 1;
IF rst OR NOT init THEN
	init := TRUE;
	FOR i := 0 TO stop DO buf[i] := in; END_FOR;
	out := in;
	i := 0;
ELSIF stop < 0 THEN
	out := in;
ELSE
	out := buf[i];
	buf[i] := in;
	i := INC1(i, N);
END_IF;

(* revision history
hm 1.10.2006		rev 1.1
	corrected error in buffer management

hm 19.1.2007		rev 1.2
	changed reset to load the value of in instead of 0

hm	27. oct. 2008	rev 1.3
	improved performance

hm	23. feb.2009	rev 1.4
	corrected an index problem

hm	23. mar. 2009	rev 1.5
	corrected non standard write to input N

*)
(*@KEY@: END_WORKSHEET *)
END_FUNCTION_BLOCK

(* ---- DELAY_4.ST ---- *)
(*@PROPERTIES_EX@
TYPE: POU
LOCALE: 0
IEC_LANGUAGE: ST
PLC_TYPE: independent
PROC_TYPE: independent
GROUP: ENGINEERING.SIGNAL_PROCESSING
*)
(*@KEY@:DESCRIPTION*)
version 1.1	19 jan 2007
programmer 	hugo
tested by	tobias

this function block delays input values by each programm cycle
after 4 cycles the in value has shifted to the out 4 and will be discarded after the next cycle
the blocks can be cascaded.
(*@KEY@:END_DESCRIPTION*)
FUNCTION_BLOCK DELAY_4

(*Group:Default*)

VAR_INPUT
	IN :	REAL;
END_VAR

VAR_OUTPUT
	OUT1 :	REAL;
	OUT2 :	REAL;
	OUT3 :	REAL;
	OUT4 :	REAL;
END_VAR

VAR
	temp :	REAL;
END_VAR

(*@KEY@: WORKSHEET
NAME: DELAY_4
IEC_LANGUAGE: ST
*)
out4 := out3;
out3 := out2;
out2 := out1;
out1 := temp;
temp := in;

(* revision history

hm 19.1.2007	rev 1.1
	added variable temp to add 1 delay  for q1

*)
(*@KEY@: END_WORKSHEET *)
END_FUNCTION_BLOCK

(* ---- DRIVER_1.ST ---- *)
(*@PROPERTIES_EX@
TYPE: POU
LOCALE: 0
IEC_LANGUAGE: ST
PLC_TYPE: independent
PROC_TYPE: independent
GROUP: ENGINEERING.AUTOMATION
*)
(*@KEY@:DESCRIPTION*)
version 1.0	2 jan 2008
programmer 	hugo
tested by	tobias

driver_1 is a multi purpose driver.
a rising edge in in sets the output high if toggle is flase. while toggle is true, a rising edge on in toggles the output Q.
if a timeout is specified the output q will be reset to false automatically after the timeout has elapsed.
a asynchronous reset and set will force the output high or low respectively.
(*@KEY@:END_DESCRIPTION*)
FUNCTION_BLOCK DRIVER_1

(*Group:Default*)

VAR_INPUT
	SET :	BOOL;
	IN :	BOOL;
	RST :	BOOL;
	TOGGLE_MODE :	BOOL;
	TIMEOUT :	TIME;
END_VAR

VAR_OUTPUT
	Q :	BOOL;
END_VAR

VAR
	off :	TON;
	edge :	BOOL;
END_VAR

(*@KEY@: WORKSHEET
NAME: DRIVER_1
IEC_LANGUAGE: ST
*)
IF off.Q THEN Q := FALSE; END_IF;
IF rst THEN
	Q := FALSE;
ELSIF set THEN
	Q := TRUE;
ELSIF IN AND NOT edge THEN
	IF toggle_mode THEN q := NOT Q; ELSE q := TRUE; END_IF;
END_IF;
edge := in;
IF timeout > t#0s THEN off(in := Q, PT := Timeout); END_IF;

(* revision history
hm	2. jan 2008		rev 1.0
	original version

*)
(*@KEY@: END_WORKSHEET *)
END_FUNCTION_BLOCK

(* ---- DRIVER_4.ST ---- *)
(*@PROPERTIES_EX@
TYPE: POU
LOCALE: 0
IEC_LANGUAGE: ST
PLC_TYPE: independent
PROC_TYPE: independent
GROUP: ENGINEERING.AUTOMATION
*)
(*@KEY@:DESCRIPTION*)
version 1.0	2 jan 2008
programmer 	hugo
tested by	tobias

driver_4 is a multi purpose driver.
a rising edge in in sets the output high if toggle is flase. while toggle is true, a rising edge on in toggles the output Q.
if a timeout is specified the output q will be reset to false automatically after the timeout has elapsed.
a asynchronous reset and set will force the output high or low respectively.
(*@KEY@:END_DESCRIPTION*)
FUNCTION_BLOCK DRIVER_4

(*Group:Default*)

VAR_INPUT
	SET :	BOOL;
	IN0 :	BOOL;
	IN1 :	BOOL;
	IN2 :	BOOL;
	IN3 :	BOOL;
	RST :	BOOL;
	TOGGLE_MODE :	BOOL;
	TIMEOUT :	TIME;
END_VAR

VAR_OUTPUT
	Q0 :	BOOL;
	Q1 :	BOOL;
	Q2 :	BOOL;
	Q3 :	BOOL;
END_VAR

VAR
	d0 :	DRIVER_1;
	d1 :	DRIVER_1;
	d2 :	DRIVER_1;
	d3 :	DRIVER_1;
END_VAR

(*@KEY@: WORKSHEET
NAME: DRIVER_4
IEC_LANGUAGE: ST
*)
D0(Set:=set, in:=in0, rst:=rst, toggle_mode:=toggle_mode, timeout:=timeout);
D1(Set:=set, in:=in1, rst:=rst, toggle_mode:=toggle_mode, timeout:=timeout);
D2(Set:=set, in:=in2, rst:=rst, toggle_mode:=toggle_mode, timeout:=timeout);
D3(Set:=set, in:=in3, rst:=rst, toggle_mode:=toggle_mode, timeout:=timeout);
Q0 := D0.Q;
Q1 := D1.Q;
Q2 := D2.Q;
Q3 := D3.Q;

(* revision history
hm	2. jan 2008		rev 1.0
	original version

*)
(*@KEY@: END_WORKSHEET *)
END_FUNCTION_BLOCK

(* ---- DRIVER_4C.ST ---- *)
(*@PROPERTIES_EX@
TYPE: POU
LOCALE: 0
IEC_LANGUAGE: ST
PLC_TYPE: independent
PROC_TYPE: independent
GROUP: ENGINEERING.AUTOMATION
*)
(*@KEY@:DESCRIPTION*)
version 1.0	23. mar. 2009
programmer 	hugo
tested by	tobias

driver_4C is a multi purpose driver.
a rising edge on in switches from S0 state S1 and the next edge to state S2 and so on.
in state S0 all outputs Q are FALSE.
The stet of the Outputs in any state S? is configurable with setup variables.
The variables S1..S5 define the states, while the sequence is terminated when a state Variable S? = 0.
The lower bits 0..3 of the state vars S? are corresponding to the Outputs Q0..Q3

(*@KEY@:END_DESCRIPTION*)
FUNCTION_BLOCK DRIVER_4C

(*Group:Default*)

VAR_INPUT
	IN :	BOOL;
	RST :	BOOL;
	TIMEOUT :	TIME;
	SX :	oscat_DRIVER_4C;
END_VAR

VAR_OUTPUT
	SN :	INT;
	Q0 :	BOOL;
	Q1 :	BOOL;
	Q2 :	BOOL;
	Q3 :	BOOL;
END_VAR

VAR
	off :	TON;
	edge :	BOOL;
END_VAR

(*@KEY@: WORKSHEET
NAME: DRIVER_4C
IEC_LANGUAGE: ST
*)
IF RST OR off.Q THEN
	SN := 0;
ELSIF IN AND NOT edge THEN
	SN := SN + 1;
	IF SN > 7 OR SX[SN] = BYTE#0 THEN SN := 0; END_IF;
END_IF;
edge := in;
IF SN > 0 THEN
	Q0 := (SX[SN] AND BYTE#1) > BYTE#0;
	Q1 := (SX[SN] AND BYTE#2) > BYTE#0;
	Q2 := (SX[SN] AND BYTE#4) > BYTE#0;
	Q3 := (SX[SN] AND BYTE#8) > BYTE#0;
ELSE
	Q0 := FALSE;
	Q1 := FALSE;
	Q2 := FALSE;
	Q3 := FALSE;
END_IF;

(* maximaum timeout *)
IF timeout > t#0s THEN off(in := SN > 0, PT := Timeout); END_IF;

(* revision history
hm	23. mar. 2009	rev 1.0
	original version

*)
(*@KEY@: END_WORKSHEET *)
END_FUNCTION_BLOCK

(* ---- ENERGY.ST ---- *)
(*@PROPERTIES_EX@
TYPE: POU
LOCALE: 0
IEC_LANGUAGE: ST
PLC_TYPE: independent
PROC_TYPE: independent
GROUP: ENGINEERING.CONVERSION
*)
(*@KEY@:DESCRIPTION*)
version 1.2	16. jan. 2010
programmer 	hugo
tested by	oscat

this function converts different energy units
any unused input can simply be left open.
different inputs connected at the same time will be added up.
(*@KEY@:END_DESCRIPTION*)
FUNCTION_BLOCK ENERGY

(*Group:Default*)

VAR_INPUT
	J :	REAL;
	C :	REAL;
	WH :	REAL;
END_VAR

VAR_OUTPUT
	YJ :	REAL;
	YC :	REAL;
	YWH :	REAL;
END_VAR

(*@KEY@: WORKSHEET
NAME: ENERGY
IEC_LANGUAGE: ST
*)
YJ := J + Wh * 3600.0 + C * 4.1868;
YC := YJ * 0.238845896627496;
YWh := YJ * 2.7777777778E-004;

(*
Arbeit, Energie, Joule* J 1 J = 1 N · m = 1 W · s = (1/3,6) E–6 kW · h = 1 kg · m2/s2
Wärmemenge Kilowattstunde kW · h 1 kW · h = 3,6 MJ = 860 kcal
Elektronvolt eV 1 eV = 160,218 92 E–21 J
Erg erg 1 erg = 1E–7 J
Kalorie calorie 1 calalorie = 4,1868 J = 1,163 E–3 W · h
Therm therm 1 therm = 105,50 · 106 J
*)

(* revision history

hm	27. mar. 2007	rev 1.0
	original version

hm	11. mar. 2009	rev 1.1
	improved code

hm 16. jan 2010	rev 1.2
	avoid the string cal in comments for codesys import bug

*)
(*@KEY@: END_WORKSHEET *)
END_FUNCTION_BLOCK

(* ---- ESR_COLLECT.ST ---- *)
(*@PROPERTIES_EX@
TYPE: POU
LOCALE: 0
IEC_LANGUAGE: ST
PLC_TYPE: independent
PROC_TYPE: independent
GROUP: OTHER
*)
(*@KEY@:DESCRIPTION*)
version 1.4	1. dec. 2009
programmer 	hugo
tested by	tobias

ESR_collect collects esr data from up to 8 esr_mon modules and stroes them in an output array.
the output pos will display the position of the last element in the array. if the array is empty, pos = -1
when to buffer is read by followon modules. pos has to be reset to -1
if the array will be full, the buffer will be refilled starting at position 0.

(*@KEY@:END_DESCRIPTION*)
FUNCTION_BLOCK ESR_COLLECT

(*Group:Default*)

VAR_INPUT
	ESR_0 :	oscat_ESR_3;
	ESR_1 :	oscat_ESR_3;
	ESR_2 :	oscat_ESR_3;
	ESR_3 :	oscat_ESR_3;
	ESR_4 :	oscat_ESR_3;
	ESR_5 :	oscat_ESR_3;
	ESR_6 :	oscat_ESR_3;
	ESR_7 :	oscat_ESR_3;
	RST :	BOOL;
END_VAR

VAR_IN_OUT
	POS :	INT;
END_VAR

VAR_OUTPUT
	ESR_OUT :	oscat_ESR_31;
END_VAR

VAR
	cnt :	INT := -1;
	max_in :	INT := 3;
	max_out :	INT := 32;
END_VAR

(*@KEY@: WORKSHEET
NAME: ESR_COLLECT
IEC_LANGUAGE: ST
*)
IF rst OR cnt < 0 THEN
	pos := -1;
ELSE
	FOR cnt := 0 TO max_in DO
	IF esr_0[cnt].typ > BYTE#0 THEN pos := INC1(pos, max_out); esr_out[pos] := esr_0[cnt]; END_IF;
	IF esr_1[cnt].typ > BYTE#0 THEN pos := INC1(pos, max_out); esr_out[pos] := esr_1[cnt]; END_IF;
	IF esr_2[cnt].typ > BYTE#0 THEN pos := INC1(pos, max_out); esr_out[pos] := esr_2[cnt]; END_IF;
	IF esr_3[cnt].typ > BYTE#0 THEN pos := INC1(pos, max_out); esr_out[pos] := esr_3[cnt]; END_IF;
	IF esr_4[cnt].typ > BYTE#0 THEN pos := INC1(pos, max_out); esr_out[pos] := esr_4[cnt]; END_IF;
	IF esr_5[cnt].typ > BYTE#0 THEN pos := INC1(pos, max_out); esr_out[pos] := esr_5[cnt]; END_IF;
	IF esr_6[cnt].typ > BYTE#0 THEN pos := INC1(pos, max_out); esr_out[pos] := esr_6[cnt]; END_IF;
	IF esr_7[cnt].typ > BYTE#0 THEN pos := INC1(pos, max_out); esr_out[pos] := esr_7[cnt]; END_IF;
   END_FOR;
END_IF;

(* revision history
hm	26.jan 2007	rev 1.0
	original version

hm	8. dec 2007	rev 1.1
	added reset input

ks	27. oct. 2008	rev 1.2
	optimized code for performance

ks	12. nov. 2009	rev 1.3
	output pos was not pointing to last value

hm	1. dec. 2009	rev 1.4
	changed pos to be I/O
	reduced output array size to 32 elements
*)
(*@KEY@: END_WORKSHEET *)
END_FUNCTION_BLOCK

(* ---- ESR_MON_B8.ST ---- *)
(*@PROPERTIES_EX@
TYPE: POU
LOCALE: 0
IEC_LANGUAGE: ST
PLC_TYPE: independent
PROC_TYPE: independent
GROUP: OTHER
*)
(*@KEY@:DESCRIPTION*)
version 1.3	1. dec. 2009
programmer 	hugo
tested by	tobias

ESR_mon_B8 monitores up to 8 binary inputs and reports changes with time stamd and adress label.
the module checks 8 inputs for a change and reports all changes with time and adress stamp to the output.
4 events maximum can be collected at once within the same cycle

(*@KEY@:END_DESCRIPTION*)
FUNCTION_BLOCK ESR_MON_B8

(*Group:Default*)

VAR_INPUT
	S0 :	BOOL;
	A0 :	oscat_STRING10;
	S1 :	BOOL;
	A1 :	oscat_STRING10;
	S2 :	BOOL;
	A2 :	oscat_STRING10;
	S3 :	BOOL;
	A3 :	oscat_STRING10;
	S4 :	BOOL;
	A4 :	oscat_STRING10;
	S5 :	BOOL;
	A5 :	oscat_STRING10;
	S6 :	BOOL;
	A6 :	oscat_STRING10;
	S7 :	BOOL;
	A7 :	oscat_STRING10;
	DT_IN :	UDINT;
END_VAR

VAR_IN_OUT
	ESR_Out :	oscat_ESR_3;
END_VAR

VAR_OUTPUT
	ESR_FLAG :	BOOL;
END_VAR

VAR
	x0 :	BOOL;
	x1 :	BOOL;
	x2 :	BOOL;
	x3 :	BOOL;
	x4 :	BOOL;
	x5 :	BOOL;
	x6 :	BOOL;
	x7 :	BOOL;
	tx :	TIME;
	cnt :	INT;
	T_PLC_MS :	T_PLC_MS;
END_VAR

(*@KEY@: WORKSHEET
NAME: ESR_MON_B8
IEC_LANGUAGE: ST
*)
(* read system timer *)
T_PLC_MS();
tx:= UDINT_TO_TIME(T_PLC_MS.T_PLC_MS);

ESR_Flag := FALSE;
esr_out[3].typ := BYTE#0;
esr_out[2].typ := BYTE#0;
esr_out[1].typ := BYTE#0;
esr_out[0].typ := BYTE#0;
cnt := 0;

(* check if inputs have chaged and fill buffer *)
IF s0 <> X0 THEN
	esr_out[cnt].typ := INT_TO_BYTE(10 + BOOL_TO_INT(s0));
	esr_out[cnt].adress := a0;
	esr_out[cnt].DS := DT_in;
	esr_out[cnt].TS := TX;
	X0 := S0;
	cnt := cnt + 1;
	esr_flag := TRUE;
END_IF;
IF s1 <> X1 THEN
	esr_out[cnt].typ := INT_TO_BYTE(10 + BOOL_TO_INT(s1));
	esr_out[cnt].adress := a1;
	esr_out[cnt].DS := DT_in;
	esr_out[cnt].TS := TX;
	X1 := S1;
	cnt := cnt + 1;
	esr_flag := TRUE;
END_IF;
IF s2 <> X2 THEN
	esr_out[cnt].typ := INT_TO_BYTE(10 + BOOL_TO_INT(s2));
	esr_out[cnt].adress := a2;
	esr_out[cnt].DS := DT_in;
	esr_out[cnt].TS := TX;
	X2 := S2;
	cnt := cnt + 1;
	esr_flag := TRUE;
END_IF;
IF s3 <> X3 THEN
	esr_out[cnt].typ := INT_TO_BYTE(10 + BOOL_TO_INT(s3));
	esr_out[cnt].adress := a3;
	esr_out[cnt].DS := DT_in;
	esr_out[cnt].TS := TX;
	X3 := S3;
	cnt := cnt + 1;
	esr_flag := TRUE;
END_IF;
IF s4 <> X4 AND cnt < 4 THEN
	esr_out[cnt].typ := INT_TO_BYTE(10 + BOOL_TO_INT(s4));
	esr_out[cnt].adress := a4;
	esr_out[cnt].DS := DT_in;
	esr_out[cnt].TS := TX;
	X4 := S4;
	cnt := cnt + 1;
	esr_flag := TRUE;
END_IF;
IF s5 <> X5  AND cnt < 4 THEN
	esr_out[cnt].typ := INT_TO_BYTE(10 + BOOL_TO_INT(s5));
	esr_out[cnt].adress := a5;
	esr_out[cnt].DS := DT_in;
	esr_out[cnt].TS := TX;
	X5 := S5;
	cnt := cnt + 1;
	esr_flag := TRUE;
END_IF;
IF s6 <> X6  AND cnt < 4 THEN
	esr_out[cnt].typ := INT_TO_BYTE(10 + BOOL_TO_INT(s6));
	esr_out[cnt].adress := a6;
	esr_out[cnt].DS := DT_in;
	esr_out[cnt].TS := TX;
	X6 := S6;
	cnt := cnt + 1;
	esr_flag := TRUE;
END_IF;
IF s7 <> X7  AND cnt < 4 THEN
	esr_out[cnt].typ := INT_TO_BYTE(10 + BOOL_TO_INT(s7));
	esr_out[cnt].adress := a7;
	esr_out[cnt].DS := DT_in;
	esr_out[cnt].TS := TX;
	X7 := S7;
	cnt := cnt + 1;
	esr_flag := TRUE;
END_IF;

(* revision history
hm	26. jan 2007	rev 1.0
	original version

hm	17. sep 2007	rev 1.1
	replaced time() with T_PLC_MS() for compatibility reasons

hm	22. oct. 2008	rev 1.2
	optimized code

hm	1.dec. 2009	rev 1.3
	changed esr_out to be I/O

*)
(*@KEY@: END_WORKSHEET *)
END_FUNCTION_BLOCK

(* ---- ESR_MON_R4.ST ---- *)
(*@PROPERTIES_EX@
TYPE: POU
LOCALE: 0
IEC_LANGUAGE: ST
PLC_TYPE: independent
PROC_TYPE: independent
GROUP: OTHER
*)
(*@KEY@:DESCRIPTION*)
version 1.4	1. dec. 2009
programmer 	hugo
tested by	tobias

ESR_mon_R4 monitores up to 4 Real inputs and reports changes with time stamd and adress label.
the module checks 4 inputs for a change of more than the specified sensitivity S and reports all changes with time and adress stamp to the output.

(*@KEY@:END_DESCRIPTION*)
FUNCTION_BLOCK ESR_MON_R4

(*Group:Default*)

VAR_INPUT
	R0 :	REAL;
	A0 :	oscat_STRING10;
	S0 :	REAL;
	R1 :	REAL;
	A1 :	oscat_STRING10;
	S1 :	REAL;
	R2 :	REAL;
	A2 :	oscat_STRING10;
	S2 :	REAL;
	R3 :	REAL;
	A3 :	oscat_STRING10;
	S3 :	REAL;
	DT_IN :	UDINT;
END_VAR

VAR_IN_OUT
	ESR_OUT :	oscat_ESR_3;
END_VAR

VAR_OUTPUT
	ESR_FLAG :	BOOL;
END_VAR

VAR
	x0 :	REAL;
	x1 :	REAL;
	x2 :	REAL;
	x3 :	REAL;
	tx :	TIME;
	cnt :	INT;
	T_PLC_MS :	T_PLC_MS;
	REAL_TO_DW :	REAL_TO_DW;
	tmp :	DWORD;
END_VAR

(*@KEY@: WORKSHEET
NAME: ESR_MON_R4
IEC_LANGUAGE: ST
*)
T_PLC_MS();
tx:= UDINT_TO_TIME(T_PLC_MS.T_PLC_MS);

ESR_Flag := FALSE;
esr_out[3].typ := BYTE#0;
esr_out[2].typ := BYTE#0;
esr_out[1].typ := BYTE#0;
esr_out[0].typ := BYTE#0;
cnt := 0;

(* check if inputs have chaged and fill buffer *)
IF differ(R0, X0, S0) THEN
    REAL_TO_DW(X:=R0);
    tmp := REAL_TO_DW.REAL_TO_DW;

	esr_out[cnt].typ := BYTE#20;
	esr_out[cnt].adress := a0;
	esr_out[cnt].DS := DT_in;
	esr_out[cnt].TS := TX;
	esr_out[cnt].data[0] := Byte_of_Dword(tmp,BYTE#0);
	esr_out[cnt].data[1] := Byte_of_Dword(tmp,BYTE#1);
	esr_out[cnt].data[2] := Byte_of_Dword(tmp,BYTE#2);
	esr_out[cnt].data[3] := Byte_of_Dword(tmp,BYTE#3);
	X0 := R0;
	cnt := cnt + 1;
	esr_flag := TRUE;
END_IF;
IF differ(R1, X1, S1) THEN
    REAL_TO_DW(X:=R1);
    tmp := REAL_TO_DW.REAL_TO_DW;

	esr_out[cnt].typ := BYTE#20;
	esr_out[cnt].adress := a1;
	esr_out[cnt].DS := DT_in;
	esr_out[cnt].TS := TX;
	esr_out[cnt].data[0] := Byte_of_Dword(tmp,BYTE#0);
	esr_out[cnt].data[1] := Byte_of_Dword(tmp,BYTE#1);
	esr_out[cnt].data[2] := Byte_of_Dword(tmp,BYTE#2);
	esr_out[cnt].data[3] := Byte_of_Dword(tmp,BYTE#3);
	X1 := R1;
	cnt := cnt + 1;
	esr_flag := TRUE;
END_IF;
IF differ(R2, X2, S2) THEN
    REAL_TO_DW(X:=R2);
    tmp := REAL_TO_DW.REAL_TO_DW;

	esr_out[cnt].typ := BYTE#20;
	esr_out[cnt].adress := a2;
	esr_out[cnt].DS := DT_in;
	esr_out[cnt].TS := TX;
	esr_out[cnt].data[0] := Byte_of_Dword(tmp,BYTE#0);
	esr_out[cnt].data[1] := Byte_of_Dword(tmp,BYTE#1);
	esr_out[cnt].data[2] := Byte_of_Dword(tmp,BYTE#2);
	esr_out[cnt].data[3] := Byte_of_Dword(tmp,BYTE#3);
	X2 := R2;
	cnt := cnt + 1;
	esr_flag := TRUE;
END_IF;
IF differ(R3, X3, S3) THEN
    REAL_TO_DW(X:=R2);
    tmp := REAL_TO_DW.REAL_TO_DW;

	esr_out[cnt].typ := BYTE#20;
	esr_out[cnt].adress := a3;
	esr_out[cnt].DS := DT_in;
	esr_out[cnt].TS := TX;
	esr_out[cnt].data[0] := Byte_of_Dword(tmp,BYTE#0);
	esr_out[cnt].data[1] := Byte_of_Dword(tmp,BYTE#1);
	esr_out[cnt].data[2] := Byte_of_Dword(tmp,BYTE#2);
	esr_out[cnt].data[3] := Byte_of_Dword(tmp,BYTE#3);
	X3 := R3;
	cnt := cnt + 1;
	esr_flag := TRUE;
END_IF;

(* revision history
hm	26. jan 2007	rev 1.0
	original version

hm	17. sep. 2007		rev 1.1
	replaced time() with T_PLC_MS() for compatibility reasons

hm	8. dec. 2007		rev 1.2
	corrected an error while esr typ would not be set

hm	16. mar. 2008		rev 1.3
	deleted wrong conversion real_to_dword

hm	1. dec 2009		rev 1.4
	changed esr_out to be I/O

*)

(*@KEY@: END_WORKSHEET *)
END_FUNCTION_BLOCK

(* ---- ESR_MON_X8.ST ---- *)
(*@PROPERTIES_EX@
TYPE: POU
LOCALE: 0
IEC_LANGUAGE: ST
PLC_TYPE: independent
PROC_TYPE: independent
GROUP: OTHER
*)
(*@KEY@:DESCRIPTION*)
version 1.2	1. dec. 2009
programmer 	hugo
tested by	tobias

ESR_MON_X8 is a status and error collector.
the module checks 8 status inputs for a change and reports up to 4 input changes with time and adress stamp to the output.
the mode can be
1 for error only
2 for error and status
3 for error, status and debug
the adress label of the 8 inputs can be configured individually.
(*@KEY@:END_DESCRIPTION*)
FUNCTION_BLOCK ESR_MON_X8

(*Group:Default*)

VAR_INPUT
	S0 :	BYTE;
	A0 :	oscat_STRING10;
	S1 :	BYTE;
	A1 :	oscat_STRING10;
	S2 :	BYTE;
	A2 :	oscat_STRING10;
	S3 :	BYTE;
	A3 :	oscat_STRING10;
	S4 :	BYTE;
	A4 :	oscat_STRING10;
	S5 :	BYTE;
	A5 :	oscat_STRING10;
	S6 :	BYTE;
	A6 :	oscat_STRING10;
	S7 :	BYTE;
	A7 :	oscat_STRING10;
	DT_IN :	UDINT;
	MODE :	BYTE := BYTE#3;
END_VAR

VAR_IN_OUT
	ESR_OUT :	oscat_ESR_3;
END_VAR

VAR_OUTPUT
	ESR_FLAG :	BOOL;
END_VAR

VAR
	x0 :	BYTE;
	x1 :	BYTE;
	x2 :	BYTE;
	x3 :	BYTE;
	x4 :	BYTE;
	x5 :	BYTE;
	x6 :	BYTE;
	x7 :	BYTE;
	tx :	TIME;
	cnt :	INT;
	status_to_ESR :	status_to_ESR;
	T_PLC_MS :	T_PLC_MS;
END_VAR

(*@KEY@: WORKSHEET
NAME: ESR_MON_X8
IEC_LANGUAGE: ST
*)
(* read system timer *)
T_PLC_MS();
tx:= UDINT_TO_TIME(T_PLC_MS.T_PLC_MS);

ESR_Flag := FALSE;
esr_out[3].typ := BYTE#0;
esr_out[2].typ := BYTE#0;
esr_out[1].typ := BYTE#0;
esr_out[0].typ := BYTE#0;
cnt := 0;

(* check if inputs have chaged and fill buffer *)
IF s0 <> X0 AND ((s0 < BYTE#100) OR (S0 > BYTE#99 AND S0 < BYTE#200 AND mode >= BYTE#2) OR (S0 > BYTE#199 AND mode = BYTE#3)) THEN

    status_to_ESR.status := s0;
    status_to_ESR.adress := a0;
    status_to_ESR.DT_in  := DT_in;
    status_to_ESR.TS     := tx;
    status_to_ESR();
    esr_out[cnt] := status_to_ESR.status_to_ESR;

	X0 := S0;
	cnt := cnt + 1;
	esr_flag := TRUE;
END_IF;
IF s1 <> X1 AND ((s1 < BYTE#100) OR (S1 > BYTE#99 AND S1 < BYTE#200 AND mode >= BYTE#2) OR (S1 > BYTE#199 AND mode = BYTE#3)) THEN

    status_to_ESR.status := s1;
    status_to_ESR.adress := a1;
    status_to_ESR.DT_in  := DT_in;
    status_to_ESR.TS     := tx;
    status_to_ESR();
    esr_out[cnt] := status_to_ESR.status_to_ESR;

	X1 := S1;
	cnt := cnt + 1;
	esr_flag := TRUE;
END_IF;
IF s2 <> X2 AND ((s2 < BYTE#100) OR (S2 > BYTE#99 AND S2 < BYTE#200 AND mode >= BYTE#2) OR (S2 > BYTE#199 AND mode = BYTE#3)) THEN

    status_to_ESR.status := s2;
    status_to_ESR.adress := a2;
    status_to_ESR.DT_in  := DT_in;
    status_to_ESR.TS     := tx;
    status_to_ESR();
    esr_out[cnt] := status_to_ESR.status_to_ESR;

	X2 := S2;
	cnt := cnt + 1;
	esr_flag := TRUE;
END_IF;
IF s3 <> X3 AND ((s3 < BYTE#100) OR (S3 > BYTE#99 AND S3 < BYTE#200 AND mode >= BYTE#2) OR (S3 > BYTE#199 AND mode = BYTE#3)) THEN

    status_to_ESR.status := s3;
    status_to_ESR.adress := a3;
    status_to_ESR.DT_in  := DT_in;
    status_to_ESR.TS     := tx;
    status_to_ESR();
    esr_out[cnt] := status_to_ESR.status_to_ESR;

	X3 := S3;
	cnt := cnt + 1;
	esr_flag := TRUE;
END_IF;
IF cnt < 4 AND s4 <> X4 AND ((s4 < BYTE#100) OR (S4 > BYTE#99 AND S4 < BYTE#200 AND mode >= BYTE#2) OR (S4 > BYTE#199 AND mode = BYTE#3)) THEN

    status_to_ESR.status := s4;
    status_to_ESR.adress := a4;
    status_to_ESR.DT_in  := DT_in;
    status_to_ESR.TS     := tx;
    status_to_ESR();
    esr_out[cnt] := status_to_ESR.status_to_ESR;

	X4 := S4;
	cnt := cnt + 1;
	esr_flag := TRUE;
END_IF;
IF cnt < 4 AND s5 <> X5 AND ((s5 < BYTE#100) OR (S5 > BYTE#99 AND S5 < BYTE#200 AND mode >= BYTE#2) OR (S5 > BYTE#199 AND mode = BYTE#3)) THEN

    status_to_ESR.status := s5;
    status_to_ESR.adress := a5;
    status_to_ESR.DT_in  := DT_in;
    status_to_ESR.TS     := tx;
    status_to_ESR();
    esr_out[cnt] := status_to_ESR.status_to_ESR;

	X5 := S5;
	cnt := cnt + 1;
	esr_flag := TRUE;
END_IF;
IF cnt < 4 AND s6 <> X6 AND ((s6 < BYTE#100) OR (S6 > BYTE#99 AND S6 < BYTE#200 AND mode >= BYTE#2) OR (S6 > BYTE#199 AND mode = BYTE#3)) THEN

    status_to_ESR.status := s6;
    status_to_ESR.adress := a6;
    status_to_ESR.DT_in  := DT_in;
    status_to_ESR.TS     := tx;
    status_to_ESR();
    esr_out[cnt] := status_to_ESR.status_to_ESR;

	X6 := S6;
	cnt := cnt + 1;
	esr_flag := TRUE;
END_IF;
IF cnt < 4 AND s7 <> X7 AND ((s7 < BYTE#100) OR (S7 > BYTE#99 AND S7 < BYTE#200 AND mode >= BYTE#2) OR (S7 > BYTE#199 AND mode = BYTE#3)) THEN

    status_to_ESR.status := s7;
    status_to_ESR.adress := a7;
    status_to_ESR.DT_in  := DT_in;
    status_to_ESR.TS     := tx;
    status_to_ESR();
    esr_out[cnt] := status_to_ESR.status_to_ESR;

	X7 := S7;
	cnt := cnt + 1;
	esr_flag := TRUE;
END_IF;

(* revision history
hm	26. jan 2007		rev 1.0
	original version

hm	17. sep 2007	rev 1.1
	replaced time() with T_PLC_MS() for compatibility reasons

hm	1. dec. 2009	rev 1.2
	changed esr_out to be I/O

*)
(*@KEY@: END_WORKSHEET *)
END_FUNCTION_BLOCK

(* ---- EVENTS.ST ---- *)
(*@PROPERTIES_EX@
TYPE: POU
LOCALE: 0
IEC_LANGUAGE: ST
PLC_TYPE: independent
PROC_TYPE: independent
GROUP: TIME_DATE
*)
(*@KEY@:DESCRIPTION*)
version 1.0	18. jan. 2010
programmer 	hugo
tested by	tobias

event checks an array with a list of events and displays the event if today is one.

(*@KEY@:END_DESCRIPTION*)
FUNCTION_BLOCK EVENTS

(*Group:Default*)

VAR_INPUT
	DATE_IN :	UDINT;
	ENA :	BOOL;
END_VAR

VAR_OUTPUT
	Y :	BOOL;
	NAME :	oscat_STRING30;
END_VAR

VAR_IN_OUT
	ELIST :	oscat_HOLIDAY_DATA_0_49;
END_VAR

VAR
	i :	INT;
	last_active :	UDINT;
	size :	INT := 49;
	day_in :	DINT;
	cyr :	INT;
	lday :	DINT;
	check :	oscat_HOLIDAY_DATA;
	y_int :	BOOL;
	name_int :	oscat_STRING30;
END_VAR

(*@KEY@: WORKSHEET
NAME: EVENTS
IEC_LANGUAGE: ST
*)
(* for performance reasons only activate once a day *)
IF last_active <> date_in THEN
	last_active := DATE_IN;
	Y_int := FALSE;
	name_int := '';
	day_in := DAY_OF_DATE(DATE_IN);
	cyr := YEAR_OF_DATE(DATE_IN);

	(* search list for events *)
	FOR i := 0 TO size DO
		check := elist[i];
		lday := DAY_OF_DATE(SET_DATE(cyr,SINT_TO_INT(check.month), SINT_TO_INT(check.day)));
		IF day_in >= lday AND day_in <= lday + SINT_TO_DINT(check.use) - DINT#1 THEN
			y_int := TRUE;
			name_int := check.name;
			EXIT;
		END_IF;
	END_FOR;
END_IF;

IF ENA THEN
	Y := y_int;
	NAME := name_int;
ELSE
	Y := FALSE;
	NAME := '';
END_IF;

(* revision history
hm  18. jan. 2011	rev 1.0
	new module

*)

(*@KEY@: END_WORKSHEET *)
END_FUNCTION_BLOCK

(* ---- FADE.ST ---- *)
(*@PROPERTIES_EX@
TYPE: POU
LOCALE: 0
IEC_LANGUAGE: ST
PLC_TYPE: independent
PROC_TYPE: independent
GROUP: ENGINEERING.SIGNAL_PROCESSING
*)
(*@KEY@:DESCRIPTION*)
version 1.3	24. jan. 2009
programmer 	oscat
tested BY	oscat

FADE is used to crossfade between the inputs IN1 and IN2. The fade_over time is specified with TF.
When F = TRUE then Y = IN2 after the time TF, and when F = FALSE then Y = IN1.
(*@KEY@:END_DESCRIPTION*)
FUNCTION_BLOCK FADE

(*Group:Default*)

VAR_INPUT
	IN1 :	REAL;
	IN2 :	REAL;
	F :	BOOL;
	TF :	TIME;
	RST :	BOOL;
END_VAR

VAR_OUTPUT
	Y :	REAL;
END_VAR

VAR
	rmx :	RMP_W;
END_VAR

(*@KEY@: WORKSHEET
NAME: FADE
IEC_LANGUAGE: ST
*)
rmx(rst := rst AND NOT F, set := rst AND F, pt := TF, up := F);
Y := (in2 - In1) / 65535.0 * _WORD_TO_REAL(rmx.out) + in1;

(* revision history
hm	26. dec 2007	rev 1.0
	original version

hm	18. oct. 2008	rev 1.1
	improved performance
	changed calls for rmp_w because rmp_w has chaged

hm	17. dec. 2008	rev 1.2
	function of input f was inverted

hm	24. jan. 2009	rev 1.3
	delted unused var FF
*)
(*@KEY@: END_WORKSHEET *)
END_FUNCTION_BLOCK

(* ---- FF_D2E.ST ---- *)
(*@PROPERTIES_EX@
TYPE: POU
LOCALE: 0
IEC_LANGUAGE: ST
PLC_TYPE: independent
PROC_TYPE: independent
GROUP: LOGIC.FF_EDGE_TRIGGERED
*)
(*@KEY@:DESCRIPTION*)
version 1.3	14. mar. 2009
programmer 	hugo
tested by	oscat

dual D-type flip flop with reset and rising clock trigger
(*@KEY@:END_DESCRIPTION*)
FUNCTION_BLOCK FF_D2E

(*Group:Default*)

VAR_INPUT
	D0 :	BOOL;
	D1 :	BOOL;
	CLK :	BOOL;
	RST :	BOOL;
END_VAR

VAR_OUTPUT
	Q0 :	BOOL;
	Q1 :	BOOL;
END_VAR

VAR
	edge :	BOOL;
END_VAR

(*@KEY@: WORKSHEET
NAME: FF_D2E
IEC_LANGUAGE: ST
*)
IF rst THEN
	Q0 := FALSE;
	Q1 := FALSE;
ELSIF clk AND NOT edge THEN
	Q0 := D0;
	Q1 := D1;
END_IF;
edge := CLK;

(* revision history
hm	25. dec 2007	rev 1.0
	original version

hm	27. dec 2007	rev 1.1
	changed code for better performance

hm	30. oct. 200	rev 1.2
	deleted unnecessary init with 0

hm	14. mar. 2009	rev 1.3
	removed double assignments

*)

(*@KEY@: END_WORKSHEET *)
END_FUNCTION_BLOCK

(* ---- FF_D4E.ST ---- *)
(*@PROPERTIES_EX@
TYPE: POU
LOCALE: 0
IEC_LANGUAGE: ST
PLC_TYPE: independent
PROC_TYPE: independent
GROUP: LOGIC.FF_EDGE_TRIGGERED
*)
(*@KEY@:DESCRIPTION*)
version 1.3	14. mar. 2009
programmer 	hugo
tested by	oscat

quad D-type flip flop with reset and rising clock trigger

(*@KEY@:END_DESCRIPTION*)
FUNCTION_BLOCK FF_D4E

(*Group:Default*)

VAR_INPUT
	D0 :	BOOL;
	D1 :	BOOL;
	D2 :	BOOL;
	D3 :	BOOL;
	CLK :	BOOL;
	RST :	BOOL;
END_VAR

VAR_OUTPUT
	Q0 :	BOOL;
	Q1 :	BOOL;
	Q2 :	BOOL;
	Q3 :	BOOL;
END_VAR

VAR
	edge :	BOOL;
END_VAR

(*@KEY@: WORKSHEET
NAME: FF_D4E
IEC_LANGUAGE: ST
*)
IF rst THEN
	Q0 := FALSE;
	Q1 := FALSE;
	Q2 := FALSE;
	Q3 := FALSE;
ELSIF clk AND NOT edge THEN
	Q0 := D0;
	Q1 := D1;
	Q2 := D2;
	Q3 := D3;
END_IF;
edge := CLK;

(* revision history
hm	4. aug 2006	rev 1.0
	original version

hm	27. dec 2007	rev 1.1
	changed code for better performance

hm	30. oct. 200	rev 1.2
	deleted unnecessary init with 0

hm	14. mar. 2009	rev 1.3
	removed double assignments

*)

(*@KEY@: END_WORKSHEET *)
END_FUNCTION_BLOCK

(* ---- FF_DRE.ST ---- *)
(*@PROPERTIES_EX@
TYPE: POU
LOCALE: 0
IEC_LANGUAGE: ST
PLC_TYPE: independent
PROC_TYPE: independent
GROUP: LOGIC.FF_EDGE_TRIGGERED
*)
(*@KEY@:DESCRIPTION*)
version 1.2	30. oct. 2008
programmer 	hugo
tested by	oscat

D-type flip flop with set, reset and rising clock trigger
(*@KEY@:END_DESCRIPTION*)
FUNCTION_BLOCK FF_DRE

(*Group:Default*)

VAR_INPUT
	SET :	BOOL;
	D :	BOOL;
	CLK :	BOOL;
	RST :	BOOL;
END_VAR

VAR_OUTPUT
	Q :	BOOL;
END_VAR

VAR
	edge :	BOOL;
END_VAR

(*@KEY@: WORKSHEET
NAME: FF_DRE
IEC_LANGUAGE: ST
*)
IF rst OR set THEN
	Q := NOT rst;
ELSIF clk AND NOT edge THEN
	Q := D;
END_IF;
edge := CLK;

(* revision history
hm	4. aug 2006		rev 1.0
	original version

hm	27. dec 2007	rev 1.1
	changed code for better performance

hm	30. oct. 2008	rev 1.2
	optimized performance
*)
(*@KEY@: END_WORKSHEET *)
END_FUNCTION_BLOCK

(* ---- FF_JKE.ST ---- *)
(*@PROPERTIES_EX@
TYPE: POU
LOCALE: 0
IEC_LANGUAGE: ST
PLC_TYPE: independent
PROC_TYPE: independent
GROUP: LOGIC.FF_EDGE_TRIGGERED
*)
(*@KEY@:DESCRIPTION*)
version 1.2	30. oct. 2008
programmer 	hugo
tested by	oscat

JK-type flip flop with set, reset and rising clock trigger
set and reset are asynchron while the FF is rising edge triggered
J=0 and K=0 and CLK >>> no action
J=1 and K=0 and CLK >>> output = 1
J=0 and K=1 and CLK >>> output = 0
J=1 and K=1 and CLK >>> toggle output
(*@KEY@:END_DESCRIPTION*)
FUNCTION_BLOCK FF_JKE

(*Group:Default*)

VAR_INPUT
	SET :	BOOL;
	J :	BOOL;
	CLK :	BOOL;
	K :	BOOL;
	RST :	BOOL;
END_VAR

VAR_OUTPUT
	Q :	BOOL;
END_VAR

VAR
	edge :	BOOL;
END_VAR

(*@KEY@: WORKSHEET
NAME: FF_JKE
IEC_LANGUAGE: ST
*)
IF rst OR set THEN
	Q := NOT rst;
ELSIF clk AND NOT edge THEN
	IF J XOR K THEN Q := J;
	ELSE Q := K XOR Q;
	END_IF;
END_IF;
edge := CLK;

(* revision history
hm	4. aug 2006		rev 1.0
	original version

hm	27. dec 2007	rev 1.1
	changed code for better performance

hm	30. oct. 2008	rev 1.2
	optimized performance
*)
(*@KEY@: END_WORKSHEET *)
END_FUNCTION_BLOCK

(* ---- FF_RSE.ST ---- *)
(*@PROPERTIES_EX@
TYPE: POU
LOCALE: 0
IEC_LANGUAGE: ST
PLC_TYPE: independent
PROC_TYPE: independent
GROUP: LOGIC.FF_EDGE_TRIGGERED
*)
(*@KEY@:DESCRIPTION*)
version 1.0	16. jul. 2008
programmer 	hugo
tested by	oscat

this is a rising edge triggered rs flip flop
a rising edge on CS sets Q = TRUE and a rising edge on CR sets Q = FALSE.
CR has priority over CS.
(*@KEY@:END_DESCRIPTION*)
FUNCTION_BLOCK FF_RSE

(*Group:Default*)

VAR_INPUT
	CS :	BOOL;
	CR :	BOOL;
	RST :	BOOL;
END_VAR

VAR_OUTPUT
	Q :	BOOL;
END_VAR

VAR
	es :	BOOL;
	er :	BOOL;
END_VAR

(*@KEY@: WORKSHEET
NAME: FF_RSE
IEC_LANGUAGE: ST
*)
IF rst THEN
	(* asynchronous reset *)
	Q := FALSE;
ELSIF CR AND NOT er THEN
	(* rising edge on CR *)
	Q := FALSE;
ELSIF CS AND NOT es THEN
	(* rising edge on CS *)
	Q := TRUE;
END_IF;

es := CS;
er := CR;

(* revision history

hm	16. jul. 2008	rev 1.0
	original version

*)
(*@KEY@: END_WORKSHEET *)
END_FUNCTION_BLOCK

(* ---- FIFO_16.ST ---- *)
(*@PROPERTIES_EX@
TYPE: POU
LOCALE: 0
IEC_LANGUAGE: ST
PLC_TYPE: independent
PROC_TYPE: independent
GROUP: LOGIC.MEMORY
*)
(*@KEY@:DESCRIPTION*)
version 2.0	24. jul. 2009
programmer 	hugo
tested by	oscat

16 Dword FIFO memory
(*@KEY@:END_DESCRIPTION*)
FUNCTION_BLOCK FIFO_16

(*Group:Default*)

VAR_INPUT
	DIN :	DWORD;
	E :	BOOL := TRUE;
	RD :	BOOL;
	WD :	BOOL;
	RST :	BOOL;
END_VAR

VAR_OUTPUT
	DOUT :	DWORD;
	EMPTY :	BOOL := TRUE;
	FULL :	BOOL;
END_VAR

VAR
	fifo :	oscat_ardw_0_15;
	pr :	INT;
	pw :	INT;
END_VAR

(*@KEY@: WORKSHEET
NAME: FIFO_16
IEC_LANGUAGE: ST
*)
IF RST THEN
	pw := pr;
	FULL := FALSE;
	EMPTY := TRUE;
	Dout := DWORD#0;
ELSIF E THEN
	IF NOT EMPTY AND RD THEN
		Dout := fifo[pr];
		pr := INC1(pr,16);
		EMPTY := pr = pw;
		FULL := FALSE;
	END_IF;
	IF NOT FULL AND WD THEN
		fifo[pw] := Din;
		pw := INC1(pw,16);
		FULL := pw = pr;
		EMPTY := FALSE;
	END_IF;
END_IF;

(* revision history

hm	4. aug. 2006	rev 1.0
	original version

hm	19. feb 2008	rev 1.1
	performance improvements

hm	17. oct. 2008	rev 1.2
	improved performance

ks	27. oct. 2008	rev 1.3
	optimized coding

hm	14. mar. 2009	rev 1.4
	removed double assignments

hm 24. jul. 2009	rev 2.0
	chaged inputs E and WR to E, WD and WR
	allow read and write in one cycle

*)

(*@KEY@: END_WORKSHEET *)
END_FUNCTION_BLOCK

(* ---- FIFO_32.ST ---- *)
(*@PROPERTIES_EX@
TYPE: POU
LOCALE: 0
IEC_LANGUAGE: ST
PLC_TYPE: independent
PROC_TYPE: independent
GROUP: LOGIC.MEMORY
*)
(*@KEY@:DESCRIPTION*)
version 2.0	24. jul. 2009
programmer 	hugo
tested by	oscat

32 Dword FIFO memory
(*@KEY@:END_DESCRIPTION*)
FUNCTION_BLOCK FIFO_32

(*Group:Default*)

VAR_INPUT
	DIN :	DWORD;
	E :	BOOL := TRUE;
	RD :	BOOL;
	WD :	BOOL;
	RST :	BOOL;
END_VAR

VAR_OUTPUT
	DOUT :	DWORD;
	EMPTY :	BOOL := TRUE;
	FULL :	BOOL;
END_VAR

VAR
	fifo :	oscat_ardw_0_31;
	pr :	INT;
	pw :	INT;
END_VAR

(*@KEY@: WORKSHEET
NAME: FIFO_32
IEC_LANGUAGE: ST
*)
IF RST THEN
	pw := pr;
	FULL := FALSE;
	EMPTY := TRUE;
	Dout := DWORD#0;
ELSIF E THEN
	IF NOT EMPTY AND RD THEN
		Dout := fifo[pr];
		pr := INC1(pr,32);
		EMPTY := pr = pw;
		FULL := FALSE;
	END_IF;
	IF NOT FULL AND WD THEN
		fifo[pw] := Din;
		pw := INC1(pw,32);
		FULL := pw = pr;
		EMPTY := FALSE;
	END_IF;
END_IF;

(* revision history
hm	4. aug. 2006	rev 1.0
	original version

hm	19. feb 2008	rev 1.1
	performance improvements

hm	17. oct. 2008	rev 1.2
	improved performance

ks	27. oct. 2008 rev 1.3
	improved code

hm	14. mar. 2009	rev 1.4
	removed double assignments

hm 24. jul. 2009	rev 2.0
	chaged inputs E and WR to E, WD and WR
	allow read and write in one cycle

*)

(*@KEY@: END_WORKSHEET *)
END_FUNCTION_BLOCK

(* ---- FLOW_CONTROL.ST ---- *)
(*@PROPERTIES_EX@
TYPE: POU
LOCALE: 0
IEC_LANGUAGE: ST
PLC_TYPE: independent
PROC_TYPE: independent
GROUP: ENGINEERING.AUTOMATION
*)
(*@KEY@:DESCRIPTION*)
version 1.0	28. jun. 2008
programmer 	hugo
tested by	oscat

FLOW_CONTROL switches a valves depending on the input in.
flow control also limits the maximum ontime of the valve and controls pressure on the output side.
(*@KEY@:END_DESCRIPTION*)
FUNCTION_BLOCK FLOW_CONTROL

(*Group:Default*)

VAR_INPUT
	IN :	BOOL;
	REQ :	BOOL;
	ENQ :	BOOL;
	RST :	BOOL := FALSE;
	T_AUTO :	TIME := T#1h;
	T_DELAY :	TIME := T#23h;
END_VAR

VAR_OUTPUT
	Q :	BOOL;
	STATUS :	BYTE;
END_VAR

VAR
	timer :	TP_1D;
END_VAR

(*@KEY@: WORKSHEET
NAME: FLOW_CONTROL
IEC_LANGUAGE: ST
*)
STATUS := BYTE#100;
IF RST THEN
	Q := FALSE;
	timer(rst := TRUE);
	timer.RST := FALSE;
	STATUS := BYTE#103;
ELSIF ENQ THEN
	IF IN THEN
		status := BYTE#101;
	END_IF;
	IF REQ THEN
		(* timer will generate a timed pulse after TP goes high *)
		timer.PT1 := T_AUTO;
		timer.PTD := T_DELAY;
		timer.IN := TRUE;
		STATUS := BYTE#102;
	END_IF;
END_IF;

(* set output and run timer *)
timer();
timer.IN := FALSE;
Q := (IN AND ENQ) OR timer.Q;

(* revision history
hm 	28. jun. 2008 	rev 1.0
	original version

*)
(*@KEY@: END_WORKSHEET *)
END_FUNCTION_BLOCK

(* ---- FLOW_CONTROL_4.ST ---- *)
(*@PROPERTIES_EX@
TYPE: POU
LOCALE: 0
IEC_LANGUAGE: ST
PLC_TYPE: independent
PROC_TYPE: independent
GROUP: ENGINEERING.AUTOMATION
*)
(*@KEY@:DESCRIPTION*)
version 1.0	19. jun 2008
programmer 	hugo
tested by	oscat

FLOW_CONTROL switches up to 4 valves depending on the 4 inputs i and generates a safety valve signal.
flow control also limits the maximum ontime of valves and controls pressure on the output side.
a diangnostic mode can automatically check all valves for operation and report errors.
anti freeze can be used to protect valves from icing during cold season´.
(*@KEY@:END_DESCRIPTION*)
FUNCTION_BLOCK FLOW_CONTROL_4

(*Group:Default*)

VAR_INPUT
	I0 :	BOOL;
	I1 :	BOOL;
	I2 :	BOOL;
	I3 :	BOOL;
	PR :	BOOL;
	ICE :	BOOL;
	DIAG :	BOOL;
	ENQ :	BOOL;
	RST :	BOOL := FALSE;
	TD_WAIT :	TIME := T#5s;
	TD_S :	TIME := T#10s;
	TD_0 :	TIME := T#10s;
END_VAR

VAR_OUTPUT
	QS :	BOOL;
	Q0 :	BOOL;
	Q1 :	BOOL;
	Q2 :	BOOL;
	Q3 :	BOOL;
	ERROR :	BOOL;
	STATUS :	BYTE;
END_VAR

VAR
	state :	INT;
	timer :	TP;
END_VAR

(*@KEY@: WORKSHEET
NAME: FLOW_CONTROL_4
IEC_LANGUAGE: ST
*)
IF RST THEN
	STATUS := BYTE#100;
	state := 0;
	error := FALSE;

ELSIF DIAG THEN
	(* diag puts pressure by opening QS for TD_wait,
	thencloses all valves and waits for td_wait, opens valve_0 and checks pressure after td_0
	if pressure is too low, an error is present.
	continue the same procedure for all valves *)
	CASE state OF
		0 : (* start diag operation *)
			(* close all valves and pressurize the system *)
			QS := TRUE;
			Q0 := FALSE;
			Q1 := FALSE;
			Q2 := FALSE;
			Q3 := FALSE;
			timer(in := TRUE, pt := TD_WAIT);
			timer.IN := FALSE;
			state := 1;
		1 : (* wait for TD_wait *)
			timer();
			IF NOT timer.Q THEN
				QS := FALSE;
				timer(in := TRUE, pt := TD_S);
				timer.IN := FALSE;
				state := 2;
			END_IF;
		2:	(* wait for safety valve pressure test *)
			timer();
			IF NOT timer.Q THEN
				IF NOT pr THEN
					(* system pressure failure *)
					ERROR := TRUE;
					STATUS := BYTE#1;
					RETURN;
				END_IF;
				timer(in := TRUE, pt := TD_0);
				timer.IN := FALSE;
				Q0 := TRUE;
				state := 3;
			END_IF;
		3:	(* wait for pressure on Q0 to hold TD_0 *)
			timer();
			IF NOT timer.Q THEN
				IF NOT pr THEN
					(* valve 0 pressure failure *)
					ERROR := TRUE;
					STATUS := BYTE#1;
					RETURN;
				END_IF;
				Q0 := FALSE;
				QS := TRUE;
			END_IF;
	END_CASE;
ELSIF ICE THEN
	(* when frost is present we close the safety valve and open all other valves to depressurize the valves *)
	QS := FALSE;
	Q0 := TRUE;
	Q1 := TRUE;
	Q2 := TRUE;
	Q3 := TRUE;
	STATUS := BYTE#110;

ELSIF NOT error AND ENQ THEN
		Q0 := I0;
		Q1 := I1;
		Q2 := I2;
		Q3 := I3;
		QS := Q0 OR Q1 OR Q2 OR Q3;
		STATUS := BYTE#100;

		(* maximum ontime check *)
ELSE
	Q0 := FALSE;
	Q1 := FALSE;
	Q2 := FALSE;
	Q3 := FALSE;
END_IF;

(* revision history
hm 	19. jun. 2008 	rev 1.0
	original version

*)
(*@KEY@: END_WORKSHEET *)
END_FUNCTION_BLOCK

(* ---- FLOW_METER.ST ---- *)
(*@PROPERTIES_EX@
TYPE: POU
LOCALE: 0
IEC_LANGUAGE: ST
PLC_TYPE: independent
PROC_TYPE: independent
GROUP: ENGINEERING.MEASUREMENTS
*)
(*@KEY@:DESCRIPTION*)
version 1.0	23. jan. 2011
programmer 	hugo
tested by	oscat

Flow meter measures flow according to gated time or pulses.
(*@KEY@:END_DESCRIPTION*)
FUNCTION_BLOCK FLOW_METER

(*Group:Default*)

VAR_INPUT
	VX :	REAL;
	E :	BOOL;
	RST :	BOOL;
	PULSE_MODE :	BOOL;
	UPDATE_TIME :	TIME := T#1s;
END_VAR

VAR_OUTPUT
	F :	REAL;
END_VAR

VAR_IN_OUT
	X :	REAL;
	Y :	UDINT;
END_VAR

VAR
	T_PLC_MS :	T_PLC_MS;
	tx :	TIME;
	tl :	TIME;
	int1 :	INTEGRATE;
	init :	BOOL;
	e_last :	BOOL;
	tmp :	INT;
	x_last :	REAL;
	y_last :	UDINT;
END_VAR

(*@KEY@: WORKSHEET
NAME: FLOW_METER
IEC_LANGUAGE: ST
*)
IF NOT init THEN	(* init on power up *)
	init := TRUE;
	tl := tx;
	x_last := X;
	y_last := Y;
	int1.K := 2.7777777777777777E-4;
END_IF;

(* run integrator *)
int1(E := NOT (RST OR PULSE_MODE) AND E, X := VX, Y := X);	(* gated operation *)
X := int1.Y;

IF RST THEN		(* reset *)
	X := 0.0;
	Y := UDINT#0;
	tl := tx;
	x_last := 0.0;
	y_last := UDINT#0;
ELSIF E AND PULSE_MODE THEN	(* check for pulse mode *)
	IF NOT e_last THEN X := X + VX; END_IF;
END_IF;
e_last := E;

(* reduce X to be less than 1 and increase Y respectively *)
IF X > 1.0 THEN
	tmp := FLOOR(X);
	Y := Y + _INT_TO_UDINT(tmp);
	X := X - INT_TO_REAL(tmp);
END_IF;

(* calculate the current flow *)
T_PLC_MS();
tx := UDINT_TO_TIME(T_PLC_MS.T_PLC_MS);
IF tx - tl >= UPDATE_TIME AND UPDATE_TIME > t#0s THEN
	F := (UDINT_TO_REAL(Y - y_last) + X - x_last) / TIME_TO_REAL(tx - tl) * 3.6E6;
	y_last := Y;
	x_last := X;
	tl := tx;
END_IF;

(* revision history
hm	23. jan. 2011	rev 1.0
	original version

*)
(*@KEY@: END_WORKSHEET *)
END_FUNCTION_BLOCK

(* ---- FT_AVG.ST ---- *)
(*@PROPERTIES_EX@
TYPE: POU
LOCALE: 0
IEC_LANGUAGE: ST
PLC_TYPE: independent
PROC_TYPE: independent
GROUP: MATHEMATICAL.FUNCTIONS
*)
(*@KEY@:DESCRIPTION*)
version 1.5	10. mar. 2009
programmer 	hugo
tested by	oscat

this function calculates the moving average over n samples from a sequential input
the input values are shifted into an N deep buffer and the avg of this buffer is diplayed at anytime on the output.
a rst will load the buffer with the current in value..

(*@KEY@:END_DESCRIPTION*)
FUNCTION_BLOCK FT_AVG

(*Group:Default*)

VAR_INPUT
	IN :	REAL;
	E :	BOOL := TRUE;
	N :	INT := INT#32;
	RST :	BOOL;
END_VAR

VAR_OUTPUT
	AVG :	REAL;
END_VAR

VAR
	buff :	delay;
	i :	INT;
	init :	BOOL;
END_VAR

(*@KEY@: WORKSHEET
NAME: FT_AVG
IEC_LANGUAGE: ST
*)
(* limit n to a max of 32 because delay can do max 32 cycles *)
buff.N := LIMIT(0, N, 32);

IF NOT init OR rst THEN
	FOR i := 1 TO N DO
		buff(in := in);
	END_FOR;
	avg := in;
	init := TRUE;
ELSIF E THEN
	buff(in := in);
	avg := avg + (in - buff.out ) / INT_TO_REAL(N);
END_IF;

(* revision history

hm	7. jan. 2007	rev 1.1
	chaged rst logic to load the buffer with the actual input value instead of 0.
	added en input to allow better control of signal flow
	added init to load the buffer with in at startup to avoid rampup at beginning.
	deleted unused variable cnt.

hm	14. jun. 2008	rev 1.2
	set default for input en = TRUE and N = 32

hm	10. oct. 2008	rev 1.3
	improved performance

hm	18. oct. 2008	rev 1.4
	changed input en to e for compatibility reasons

hm	10. mar. 2009	rev 1.5
	added type conversion for compatibility reasons

*)
(*@KEY@: END_WORKSHEET *)
END_FUNCTION_BLOCK

(* ---- FT_DERIV.ST ---- *)
(*@PROPERTIES_EX@
TYPE: POU
LOCALE: 0
IEC_LANGUAGE: ST
PLC_TYPE: independent
PROC_TYPE: independent
GROUP: ENGINEERING.CONTROL
*)
(*@KEY@:DESCRIPTION*)
version 1.5	11. mar. 2009
programmer 	hugo
tested by	oscat

FT_deriv calculates the derivate over the signal "in" with Faktor "K".
a run input enables or stops the calculation, if left unconnected its true and therfore the calculation is executed.
if K is not specified the default is 1.

(*@KEY@:END_DESCRIPTION*)
FUNCTION_BLOCK FT_DERIV

(*Group:Default*)

VAR_INPUT
	IN :	REAL;
	K :	REAL := 1.0;
	RUN :	BOOL := TRUE;
END_VAR

VAR_OUTPUT
	OUT :	REAL;
END_VAR

VAR
	old :	REAL;
	tx :	UDINT;
	last :	UDINT;
	init :	BOOL;
	tc :	REAL;
	T_PLC_US :	T_PLC_US;
END_VAR

(*@KEY@: WORKSHEET
NAME: FT_DERIV
IEC_LANGUAGE: ST
*)
(* read system time *)
T_PLC_US();
tx:= T_PLC_US.T_PLC_US;
tc := UDINT_TO_REAL(tx - last);

(* init on firsat startup *)
IF NOT init THEN
	init := TRUE;
	old := in;
ELSIF run AND tc > 0.0 THEN
	out := (in - old) / tc * 1000000.0 * K;
	old := in;
ELSE
	out := 0.0;
END_IF;

last := tx;

(*
hm 3.1.2007			rev 1.1
	added init code for startup
	set the default for K to 1

hm	15. sep 2007	rev 1.2
	replaced Time() with T_PLC_US for compatibility and performance reasons
	increased accuracy and work in microseconds internally

hm 29 oct 2007	rev 1.3
	prohibit calculation when tx - last = 0 to avoid division by 0 and increase accuracy on fast systems

hm	6. nov. 2008	rev 1.4
	improved performance

hm	11. mar. 2009	rev 1.5
	inproved code
*)

(* read system time *)
T_PLC_US();
tx:= T_PLC_US.T_PLC_US;

(* init on firsat startup *)
IF NOT init THEN
	init := TRUE;
ELSIF run AND tx - last > UDINT#0 THEN
	out := (in - old) / UDINT_TO_REAL(tx - last) * 1000000.0 * K;
ELSE
	out := 0.0;
END_IF;
old := in;
last := tx;

(*
hm 3.1.2007			rev 1.1
	added init code for startup
	set the default for K to 1

hm	15. sep 2007	rev 1.2
	replaced Time() with T_PLC_US for compatibility and performance reasons
	increased accuracy and work in microseconds internally

hm 29 oct 2007	rev 1.3
	prohibit calculation when tx - last = 0 to avoid division by 0 and increase accuracy on fast systems

hm	3. nov. 2008	rev 1.4
	improved performance
*)
(*@KEY@: END_WORKSHEET *)
END_FUNCTION_BLOCK

(* ---- FT_IMP.ST ---- *)
(*@PROPERTIES_EX@
TYPE: POU
LOCALE: 0
IEC_LANGUAGE: ST
PLC_TYPE: independent
PROC_TYPE: independent
GROUP: ENGINEERING.CONTROL
*)
(*@KEY@:DESCRIPTION*)
version 1.1	3 Jan 2007
programmer 	hugo
tested by	tobias

FT_IMP is 	an impulse filter (high pass filter) with the time T and factor K.
(*@KEY@:END_DESCRIPTION*)
FUNCTION_BLOCK FT_IMP

(*Group:Default*)

VAR_INPUT
	IN :	REAL;
	T :	TIME;
	K :	REAL := 1.0;
END_VAR

VAR_OUTPUT
	OUT :	REAL;
END_VAR

VAR
	t1 :	FT_PT1;
END_VAR

(*@KEY@: WORKSHEET
NAME: FT_IMP
IEC_LANGUAGE: ST
*)
T1(in:= in, T:=T);
out := (in - t1.out) * K;

(*
hm 3.1.2007	rev 1.1
	added factor K

*)
(*@KEY@: END_WORKSHEET *)
END_FUNCTION_BLOCK

(* ---- FT_INT.ST ---- *)
(*@PROPERTIES_EX@
TYPE: POU
LOCALE: 0
IEC_LANGUAGE: ST
PLC_TYPE: independent
PROC_TYPE: independent
GROUP: ENGINEERING.CONTROL
*)
(*@KEY@:DESCRIPTION*)
version 2.2	10. mar. 2009
programmer 	hugo
tested by	oscat

FT_int is an integrator with input IN and factor K.
integration is only done while run = true, if run is false integration is stopped and the out remains at the last value.
if run is left unconnected, run is considered true by the function block.
the output ET will display the total integration time from last reset.
the out_min and out_max values can be set to ,imit the output value range.
the default for K is 1.
(*@KEY@:END_DESCRIPTION*)
FUNCTION_BLOCK FT_INT

(*Group:Default*)

VAR_INPUT
	IN :	REAL;
	K :	REAL := 1.0;
	RUN :	BOOL := TRUE;
	RST :	BOOL;
	OUT_MIN :	REAL := REAL#-1.0E-37;
	OUT_MAX :	REAL := REAL#1.0E37;
END_VAR

VAR_OUTPUT
	OUT :	REAL;
	LIM :	BOOL;
END_VAR

VAR
	INTEG :	INTEGRATE;
END_VAR

(*@KEY@: WORKSHEET
NAME: FT_INT
IEC_LANGUAGE: ST
*)
IF rst THEN
	out := 0.0;
ELSE
	integ(X := IN, E := RUN, K := K, Y := out);
	out := integ.Y;
END_IF;

(* limit the outputs *)
IF out >= OUT_MAX THEN
	out := out_max;
	LIM := TRUE;
ELSIF out <= out_min THEN
	out := out_min;
	lim := TRUE;
ELSE
	lim := FALSE;
END_IF;

(*
hm 13.12.2006	rev 1.1
	changed to "trapezregel" which increases accuracy
	before out := out + in * time new: out := out + (in + in_last) / 2 * time

hm 15.1.2007		rev 1.2
	added default for k to be 1.

hm	15.9.2007		rev 1.3
	replaced time() with T_PLC_US for compatibility and performance reason
	increased internal accuracy to microseconds

hm 29. oct 2007		rev 1.4
	changed code so int will not be called is time difference is 0 to increase accuracy on systems
	with cycle times below 1ms

hm	2. dec 2007	 	rev 1.5
	changed code for better performance

hm	5. jan 2008		rev 1.6
	further improvements in performance

hm	8. feb 2008		rev 1.7
	deleted limits +/- 1000 now limit is the range of real
	added variables out1 and out2 to extend the resolution
	corrected an error with elapsed time
	deleted unusfull output ET

hm	13. mar 2008	rev 1.8
	changed preset value out_min to -1e37.
	stop integrator at the limits.

hm	16. mar 2008	rev 1.9
	added type conversion to avoid warning under codesys 3.0

hm	2. jun. 2008	rev 2.0
	rewritten with clear code
	limits can now be set without run

hm	3. nov. 2008	rev 2.1
	optimized code using INTEGRATE and LIMX

hm	10. mar. 2009	rev 2.2
	removed nested comments
*)
(*@KEY@: END_WORKSHEET *)
END_FUNCTION_BLOCK

(* ---- FT_INT2.ST ---- *)
(*@PROPERTIES_EX@
TYPE: POU
LOCALE: 0
IEC_LANGUAGE: ST
PLC_TYPE: independent
PROC_TYPE: independent
GROUP: ENGINEERING.CONTROL
*)
(*@KEY@:DESCRIPTION*)
version 1.2	11. mar. 2009
programmer 	hugo
tested by	oscat

FT_int2 is an integrator with input IN and factor K.
integration is only done while run = true, if run is false integration is stopped and the out remains at the last value.
if run is left unconnected, run is considered true by the function block.
the out_min and out_max values can be set to ,imit the output value range.
the default for K is 1.
FT_INT2 has double presision accuracy (14 digits).
(*@KEY@:END_DESCRIPTION*)
FUNCTION_BLOCK FT_INT2

(*Group:Default*)

VAR_INPUT
	IN :	REAL;
	K :	REAL := 1.0;
	RUN :	BOOL := TRUE;
	RST :	BOOL;
	OUT_MIN :	REAL := REAL#-1.0E-37;
	OUT_MAX :	REAL := REAL#1.0E37;
END_VAR

VAR_OUTPUT
	OUT :	REAL;
	LIM :	BOOL;
END_VAR

VAR
	integ :	INTEGRATE;
	ix :	REAL;
	val :	REAL2;
	R2_ADD :	R2_ADD;
	R2_SET :	R2_SET;
END_VAR

(*@KEY@: WORKSHEET
NAME: FT_INT2
IEC_LANGUAGE: ST
*)
IF RST THEN
	R2_SET(X:=0.0);
	val:=R2_SET.R2_SET;
	out := 0.0;
ELSE
	integ(X := IN, E := RUN, K := K, Y := ix);
	ix := integ.Y;
	R2_ADD(X:=val,Y:=ix);
	val:=R2_ADD.R2_ADD;
	ix := 0.0;
	OUT := val.RX;
END_IF;

(* check output for limits *)
IF out > OUT_MIN AND out < OUT_MAX THEN
	LIM := FALSE;
ELSE
	OUT := LIMIT(OUT_MIN, OUT, OUT_MAX);
	R2_SET(X:=OUT);
	val:=R2_SET.R2_SET;
	LIM := TRUE;
END_IF;

(*	revision history
hm	2. jun. 2008	rev 1.0
	original version

hm	5. nov. 2008	rev 1.1
	rewritten code using integrate

hm	11. mar. 2009	rev 1.2
	real constants updated to new systax using dot

*)
(*@KEY@: END_WORKSHEET *)
END_FUNCTION_BLOCK

(* ---- FT_MIN_MAX.ST ---- *)
(*@PROPERTIES_EX@
TYPE: POU
LOCALE: 0
IEC_LANGUAGE: ST
PLC_TYPE: independent
PROC_TYPE: independent
GROUP: MATHEMATICAL.FUNCTIONS
*)
(*@KEY@:DESCRIPTION*)
version 1.0	1 sep 2006
programmer 	hugo
tested by	tobias

this function block stores the min and max value of an input signal.
when rst is true the mn and mx outputs are set to the in value.
when a rst is never active the function autoresets to the in value at startup.
since the input might not be present at first cycle the mn and mx are set during second cycle.
(*@KEY@:END_DESCRIPTION*)
FUNCTION_BLOCK FT_MIN_MAX

(*Group:Default*)

VAR_INPUT
	IN :	REAL;
	RST :	BOOL;
END_VAR

VAR_OUTPUT
	MX :	REAL;
	MN :	REAL;
END_VAR

VAR
	init :	BOOL;
END_VAR

(*@KEY@: WORKSHEET
NAME: FT_MIN_MAX
IEC_LANGUAGE: ST
*)
IF (rst = TRUE) OR (init = FALSE) THEN
  mn := in;
  mx := in;
  init := TRUE;
ELSIF (in < mn) THEN
  mn := in;
ELSIF (in > mx) THEN
  mx := in;
END_IF;
(*@KEY@: END_WORKSHEET *)
END_FUNCTION_BLOCK

(* ---- FT_PD.ST ---- *)
(*@PROPERTIES_EX@
TYPE: POU
LOCALE: 0
IEC_LANGUAGE: ST
PLC_TYPE: independent
PROC_TYPE: independent
GROUP: ENGINEERING.CONTROL
*)
(*@KEY@:DESCRIPTION*)
version 1.0	3. jun 2008
programmer 	hugo
tested by	tobias

FT_PD is a PD controller.
The PD controller works according to the fomula Y = KP *(IN + DERIV(e) ).
(*@KEY@:END_DESCRIPTION*)
FUNCTION_BLOCK FT_PD

(*Group:Default*)

VAR_INPUT
	IN :	REAL;
	KP :	REAL := 1.0;
	TV :	REAL := 1.0;
END_VAR

VAR_OUTPUT
	Y :	REAL;
END_VAR

VAR
	diff :	FT_DERIV;
END_VAR

(*@KEY@: WORKSHEET
NAME: FT_PD
IEC_LANGUAGE: ST
*)
(* run differentiator *)
diff(IN := IN, K := TV);

(* combine both values *)
Y := KP * (diff.out + IN);

(* revision history
hm 	3. jun. 2008 	rev 1.0
	original version

*)
(*@KEY@: END_WORKSHEET *)
END_FUNCTION_BLOCK

(* ---- FT_PDT1.ST ---- *)
(*@PROPERTIES_EX@
TYPE: POU
LOCALE: 0
IEC_LANGUAGE: ST
PLC_TYPE: independent
PROC_TYPE: independent
GROUP: ENGINEERING.CONTROL
*)
(*@KEY@:DESCRIPTION*)
version 1.0	3. jun 2008
programmer 	hugo
tested by	tobias

FT_PD is a PD controller.
The PD controller works according to the fomula Y = KP *(IN + DERIV(e) ).
(*@KEY@:END_DESCRIPTION*)
FUNCTION_BLOCK FT_PDT1

(*Group:Default*)

VAR_INPUT
	IN :	REAL;
	KP :	REAL := 1.0;
	TV :	REAL := 1.0;
	T1 :	REAL := 1.0;
END_VAR

VAR_OUTPUT
	Y :	REAL;
END_VAR

VAR
	diff :	FT_DERIV;
	TP :	FT_PT1;
END_VAR

(*@KEY@: WORKSHEET
NAME: FT_PDT1
IEC_LANGUAGE: ST
*)
(* run differentiator *)
diff(IN := IN, K := TV);

(* Run PT1 filter *)
tp(in := diff.out, T := REAL_TO_TIME(T1));

(* combine both values *)
Y := KP * (tp.out + IN);

(* revision history
hm 	3. jun. 2008 	rev 1.0
	original version

*)
(*@KEY@: END_WORKSHEET *)
END_FUNCTION_BLOCK

(* ---- FT_PI.ST ---- *)
(*@PROPERTIES_EX@
TYPE: POU
LOCALE: 0
IEC_LANGUAGE: ST
PLC_TYPE: independent
PROC_TYPE: independent
GROUP: ENGINEERING.CONTROL
*)
(*@KEY@:DESCRIPTION*)
version 2.0	3. jun 2008
programmer 	hugo
tested by	tobias

FT_PI is a PI controller.
The PID controller works according to the fomula Y = IN *(KP+ KI * INTEG(e) ).
a rst will reset the integrator to 0
ilim_h and iLim_l set the possible output range of the internal integrator.
the output flags lim will signal that the output limits are active.

default values for KP = 1, KI = 1, ILIM_L = -1E37, iLIM_H = +1E38.
(*@KEY@:END_DESCRIPTION*)
FUNCTION_BLOCK FT_PI

(*Group:Default*)

VAR_INPUT
	IN :	REAL;
	KP :	REAL := 1.0;
	KI :	REAL := 1.0;
	ILIM_L :	REAL := -1.0E38;
	ILIM_H :	REAL := 1.0E38;
	IEN :	BOOL := TRUE;
	RST :	BOOL := FALSE;
END_VAR

VAR_OUTPUT
	Y :	REAL;
	LIM :	BOOL;
END_VAR

VAR
	integ :	FT_INT;
END_VAR

(*@KEY@: WORKSHEET
NAME: FT_PI
IEC_LANGUAGE: ST
*)
(* run integrator *)
integ(IN := IN, K := KI, RUN := IEN, RST := RST, OUT_MIN := ILIM_L, OUT_MAX := ILIM_H);
(* check if integrator has reached its limits and set overflow *)
LIM := integ.LIM;
Y := KP * IN + integ.Out;

(* revision history
hm 	3. jun. 2008 	rev 2.0
	original version

*)
(*@KEY@: END_WORKSHEET *)
END_FUNCTION_BLOCK

(* ---- FT_PID.ST ---- *)
(*@PROPERTIES_EX@
TYPE: POU
LOCALE: 0
IEC_LANGUAGE: ST
PLC_TYPE: independent
PROC_TYPE: independent
GROUP: ENGINEERING.CONTROL
*)
(*@KEY@:DESCRIPTION*)
version 2.1	11. mar. 2009
programmer 	hugo
tested by	tobias

FT_PI is a PI controller.
The PID controller works according to the fomula Y = IN *(KP+ KI * INTEG(e) ).
a rst will reset the integrator to 0
ilim_h and iLim_l set the possible output range of the internal integrator.
the output flags lim will signal that the output limits are active.

default values for KP = 1, KI = 1, ILIM_L = -1E37, iLIM_H = +1E38.
(*@KEY@:END_DESCRIPTION*)
FUNCTION_BLOCK FT_PID

(*Group:Default*)

VAR_INPUT
	IN :	REAL;
	KP :	REAL := 1.0;
	TN :	REAL := 1.0;
	TV :	REAL := 1.0;
	ILIM_L :	REAL := -1.0E38;
	ILIM_H :	REAL := 1.0E38;
	IEN :	BOOL := TRUE;
	RST :	BOOL := FALSE;
END_VAR

VAR_OUTPUT
	Y :	REAL;
	LIM :	BOOL;
END_VAR

VAR
	integ :	FT_INT;
	diff :	FT_DERIV;
END_VAR

(*@KEY@: WORKSHEET
NAME: FT_PID
IEC_LANGUAGE: ST
*)
(* run integrator only if TN > 0 *)
IF TN > 0.0 THEN
	integ(IN := IN, K := 1.0 / TN, RUN := IEN, RST := RST, OUT_MIN := ILIM_L, OUT_MAX := ILIM_H);
ELSE
	integ(RST := FALSE);
END_IF;

(* run differentiator *)
diff(IN := IN, K := TV);

(* combine both values *)
Y := KP * (integ.Out + diff.out + IN);

(* check if integrator has reached its limits and set overflow *)
LIM := integ.LIM;

(* revision history
hm 3. jun. 2008 	rev 2.0
	original version

hm	11. mar. 2009	rev 2.1
	real constants updated to new systax using dot

*)
(*@KEY@: END_WORKSHEET *)
END_FUNCTION_BLOCK

(* ---- FT_PIDW.ST ---- *)
(*@PROPERTIES_EX@
TYPE: POU
LOCALE: 0
IEC_LANGUAGE: ST
PLC_TYPE: independent
PROC_TYPE: independent
GROUP: ENGINEERING.CONTROL
*)
(*@KEY@:DESCRIPTION*)
version 1.2	11. mar. 2009
programmer 	hugo
tested by	oscat

FT_PIDW is a PID controller with dynamic wind_up reset.
The PID controller works according to the fomula Y = KP *(IN + KI * INTEG(e) + DERIV(e) ).
a rst will reset the integrator to 0
lim_h and Lim_l set the possible output range of the internal integrator.
the output flags lim will signal that the output limits are active.

default values for KP = 1, KI = 1, ILIM_L = -1E37, iLIM_H = +1E38.
(*@KEY@:END_DESCRIPTION*)
FUNCTION_BLOCK FT_PIDW

(*Group:Default*)

VAR_INPUT
	IN :	REAL;
	KP :	REAL := 1.0;
	TN :	REAL := 1.0;
	TV :	REAL := 1.0;
	LIM_L :	REAL := -1.0E38;
	LIM_H :	REAL := 1.0E38;
	RST :	BOOL := FALSE;
END_VAR

VAR_OUTPUT
	Y :	REAL;
	LIM :	BOOL;
END_VAR

VAR
	integ :	INTEGRATE;
	diff :	FT_DERIV;
	YI :	REAL;
END_VAR

(*@KEY@: WORKSHEET
NAME: FT_PIDW
IEC_LANGUAGE: ST
*)
(* run the integrator *)
IF tn = 0.0 OR rst THEN
	integ(E := FALSE, Y := YI);
	YI := integ.Y;
	YI := 0.0;
ELSE
	integ(X := IN, K := 1.0 / TN, E := NOT LIM, Y := YI);
	YI := integ.Y;
END_IF;

(* add up integrator and linear part *)
Y := KP * (IN + YI);

(* run differentiator *)
diff(IN := IN, K := TV);

(* set lim before differentiator is added to stop integrator if necessary *)
IF Y > LIM_L AND Y < LIM_H THEN
	LIM := FALSE;
ELSE
	LIM := TRUE;
END_IF;

(* add differential part and limit output Y *)

Y := LIMIT(LIM_L, Y + KP * diff.out, LIM_H);

(* revision history
hm 3. jun. 2008 	rev 1.0
	original version

hm	5. nov. 2008	rev 1.1
	changed code to use integrate

hm	11. mar. 2009	rev 1.2
	real constants updated to new systax using dot

*)
(*@KEY@: END_WORKSHEET *)
END_FUNCTION_BLOCK

(* ---- FT_PIDWL.ST ---- *)
(*@PROPERTIES_EX@
TYPE: POU
LOCALE: 0
IEC_LANGUAGE: ST
PLC_TYPE: independent
PROC_TYPE: independent
GROUP: ENGINEERING.CONTROL
*)
(*@KEY@:DESCRIPTION*)
version 1.3	13. nov. 2009
programmer 	hugo
tested by	tobias

FT_PIDWL is a PID controller with dynamic wind_up reset.
The PID controller works according to the fomula Y = KP *(IN + KI * INTEG(e) + DERIV(e) ).
a rst will reset the integrator to 0
lim_h and Lim_l set the possible output range of the internal integrator.
the output flags lim will signal that the output limits are active.

default values for KP = 1, KI = 1, ILIM_L = -1E37, iLIM_H = +1E38.
(*@KEY@:END_DESCRIPTION*)
FUNCTION_BLOCK FT_PIDWL

(*Group:Default*)

VAR_INPUT
	IN :	REAL;
	KP :	REAL := 1.0;
	TN :	REAL := 1.0;
	TV :	REAL := 1.0;
	LIM_L :	REAL := -1.0E38;
	LIM_H :	REAL := 1.0E38;
	RST :	BOOL;
END_VAR

VAR_OUTPUT
	Y :	REAL;
	LIM :	BOOL;
END_VAR

VAR
	piwl :	FT_PIWL;
	diff :	FT_DERIV;
END_VAR

(*@KEY@: WORKSHEET
NAME: FT_PIDWL
IEC_LANGUAGE: ST
*)
(* if rst then *)
IF rst THEN
	piwl(rst := TRUE);
	piwl.RST := FALSE;
ELSE
	(* run PIWL controller first *)
	(* we need to check if TN = 0 and do alternative calls *)
	IF TN = 0.0 THEN
		piwl(in := IN * KP, KP := 1.0, KI := 0.0, LIM_L := LIM_L, LIM_H := LIM_H);
	ELSE
		piwl(in := IN * KP, KP := 1.0, KI := 1.0 / TN, LIM_L := LIM_L, LIM_H := LIM_H);
	END_IF;

	(* run differentiator and add_to_output *)
	diff(IN := IN, K := KP * TV);
	Y := piwl.Y + diff.out;

	(* limit the output *)
	IF Y < LIM_L THEN
		LIM := TRUE;
		Y := LIM_L;
	ELSIF Y > LIM_H THEN
		LIM := TRUE;
		Y := LIM_H;
	ELSE
		LIM := FALSE;
	END_IF;
END_IF;

(* revision history
hm 13. jun. 2008 	rev 1.0
	original version

hm	25. jan 2008	rev 1.1
	multiply differential part with KP

hm	11. mar. 2009	rev 1.2
	real constants updated to new systax using dot

hm	13. nov. 2009	rev 1.3
	fixed code for negative KP

*)
(*@KEY@: END_WORKSHEET *)
END_FUNCTION_BLOCK

(* ---- FT_PIW.ST ---- *)
(*@PROPERTIES_EX@
TYPE: POU
LOCALE: 0
IEC_LANGUAGE: ST
PLC_TYPE: independent
PROC_TYPE: independent
GROUP: ENGINEERING.CONTROL
*)
(*@KEY@:DESCRIPTION*)
version 1.0	3. jun 2008
programmer 	hugo
tested by	tobias

FT_PI is a PI controller.
The PID controller works according to the fomula Y = IN *(KP+ KI * INTEG(e) ).
a rst will reset the integrator to 0
ilim_h and iLim_l set the possible output range of the internal integrator.
the output flags lim will signal that the output limits are active.

default values for KP = 1, KI = 1, ILIM_L = -1E37, iLIM_H = +1E38.
(*@KEY@:END_DESCRIPTION*)
FUNCTION_BLOCK FT_PIW

(*Group:Default*)

VAR_INPUT
	IN :	REAL;
	KP :	REAL := 1.0;
	KI :	REAL := 1.0;
	LIM_L :	REAL := -1.0E38;
	LIM_H :	REAL := 1.0E38;
	RST :	BOOL := FALSE;
END_VAR

VAR_OUTPUT
	Y :	REAL;
	LIM :	BOOL;
END_VAR

VAR
	integ :	FT_INT;
END_VAR

(*@KEY@: WORKSHEET
NAME: FT_PIW
IEC_LANGUAGE: ST
*)
(* run integrator *)
integ(IN := IN, K := KI, RUN := NOT LIM, RST := RST);

(* set output value *)
Y := KP * IN + integ.Out;

(* check for limits *)
IF Y < LIM_L THEN
	Y := LIM_L;
	LIM := TRUE;
ELSIF Y > LIM_H THEN
	Y := LIM_H;
	LIM := TRUE;
ELSE
	LIM := FALSE;
END_IF;

(* revision history
hm 	3. jun. 2008 	rev 1.0
	original version

*)
(*@KEY@: END_WORKSHEET *)
END_FUNCTION_BLOCK

(* ---- FT_PIWL.ST ---- *)
(*@PROPERTIES_EX@
TYPE: POU
LOCALE: 0
IEC_LANGUAGE: ST
PLC_TYPE: independent
PROC_TYPE: independent
GROUP: ENGINEERING.CONTROL
*)
(*@KEY@:DESCRIPTION*)
version 1.3	11. mar. 2009
programmer 	hugo
tested by	oscat

FT_PIWL is a PI controller.
The PID controller works according to the fomula Y = IN *(KP+ KI * INTEG(e) ).
a rst will reset the integrator to 0
lim_h and Lim_l set the possible output range of the controller.
the output flag lim will signal that the output limits are active.
the integrator ist equipped with anti wind-up circuitry which limits trhe total output ranke to lim_l and lim_h

default values for KP = 1, KI = 1, ILIM_L = -1E37, iLIM_H = +1E38.

(*@KEY@:END_DESCRIPTION*)
FUNCTION_BLOCK FT_PIWL

(*Group:Default*)

VAR_INPUT
	IN :	REAL;
	KP :	REAL := 1.0;
	KI :	REAL := 1.0;
	LIM_L :	REAL := -1.0E38;
	LIM_H :	REAL := 1.0E38;
	RST :	BOOL;
END_VAR

VAR_OUTPUT
	Y :	REAL;
	LIM :	BOOL;
END_VAR

VAR
	init :	BOOL;
	tx :	UDINT;
	tc :	REAL;
	t_last :	UDINT;
	in_last :	REAL;
	i :	REAL;
	p :	REAL;
	T_PLC_US :	T_PLC_US;
END_VAR

(*@KEY@: WORKSHEET
NAME: FT_PIWL
IEC_LANGUAGE: ST
*)
(* initialize at power_up *)
IF NOT init OR RST THEN
	init := TRUE;
	in_last := in;
	T_PLC_US();
	t_last := T_PLC_US.T_PLC_US;
	i := 0.0;
	tc := 0.0;
ELSE
	(* read last cycle time in Microseconds *)
	T_PLC_US();
	tx := T_PLC_US.T_PLC_US;
	tc := UDINT_TO_REAL(tx - t_last);
	t_last := tx;

	(* calculate proportional part *)
	p := KP * IN;

	(* run integrator *)
	i := (IN + in_last) * 5.0E-7 * KI * tc + i;
	in_last := IN;

	(* calculate output Y *)
	Y := p + i;

	(* check output for limits *)
	IF Y >= LIM_H THEN
		Y := LIM_H;
		IF ki <> 0.0 THEN
			i := LIM_H - p;
		ELSE
			i := 0.0;
		END_IF;
		LIM := TRUE;
	ELSIF Y <= LIM_L THEN
		Y := LIM_L;
		IF ki <> 0.0 THEN
			i := LIM_L - p;
		ELSE
			i := 0.0;
		END_IF;
		LIM := TRUE;
	ELSE
		LIM := FALSE;
	END_IF;
END_IF;

(* revision history
hm 13. jun. 2008 	rev 1.0
	original version

hm	27. oct. 2008	rev 1.1
	integrator will not be adjusted when ki = 0

hm	25. jan 2009	rev 1.2
	module will also work with negative K

hm	11. mar. 2009	rev 1.3
	real constants updated to new systax using dot

*)
(*@KEY@: END_WORKSHEET *)
END_FUNCTION_BLOCK
